DATA_BLOCK "DB_ALARM"   // DB100
{ S7_Optimized_Access := 'FALSE' }
VERSION : 0.1
   VAR
      ALARM : Struct
         ALARM_GLOBAL : Bool;   // globální alarm
         HERMA_ERROR : Bool;
         ALARM_2 : Bool;
         ALARM_3 : Bool;
         ALARM_4 : Bool;
         ALARM_5 : Bool;
         air : Bool;   // nedostatečný tlak vzduchu
         ALARM_7 : Bool;
         ALARM_8 : Bool;
         ALARM_9 : Bool;
         ALARM_10 : Bool;
         ALARM_11 : Bool;
         ALARM_12 : Bool;
         ALARM_13 : Bool;
         ALARM_14 : Bool;
         vypadek_safety_karty : Bool;
      END_STRUCT;
      WRONG : Struct
         NENI_INICIALIZACE : Bool;
         WRONG_global : Bool;
         dvere_L_tevreny : Bool;
         dvere_P_otevreny : Bool;
         WRONG_4 : Bool;
         WRONG_5 : Bool;
         WRONG_6 : Bool;
         WRONG_7 : Bool;
         WRONG_8 : Bool;
         WRONG_9 : Bool;
         WRONG_10 : Bool;
         WRONG_11 : Bool;
         WRONG_12 : Bool;
         WRONG_13 : Bool;
         rop_glob_warning : Bool;
         rop_active_autocale : Bool;
      END_STRUCT;
      OP0 : Struct
         ALARM : Struct
            DOOR_ERROR : Bool;
            ALARM_1 : Bool;
            ALARM_2 : Bool;
            ALARM_3 : Bool;
            ALARM_4 : Bool;
            ALARM_5 : Bool;
            ALARM_6 : Bool;
            ALARM_7 : Bool;
            ALARM_8 : Bool;
            ALARM_9 : Bool;
            ALARM_10 : Bool;
            ALARM_11 : Bool;
            ALARM_12 : Bool;
            ALARM_13 : Bool;
            ALARM_14 : Bool;
            ALARM_15 : Bool;
         END_STRUCT;
         WRONG : Struct
            WRONG_0 : Bool;
            WRONG_1 : Bool;
            WRONG_2 : Bool;
            WRONG_3 : Bool;
            WRONG_4 : Bool;
            WRONG_5 : Bool;
            WRONG_6 : Bool;
            WRONG_7 : Bool;
            WRONG_8 : Bool;
            WRONG_9 : Bool;
            WRONG_10 : Bool;
            WRONG_11 : Bool;
            WRONG_12 : Bool;
            WRONG_13 : Bool;
            WRONG_14 : Bool;
            WRONG_15 : Bool;
         END_STRUCT;
         M_0 : Int;
         M_1 : Int;
         M_2 : Int;
         M_3 : Int;
         M_4 : Int;
         M_5 : Int;
         M_6 : Int;
         M_7 : Int;
         M_8 : Int;
         M_9 : Int;
         M_10 : Int;
         M_11 : Int;
         M_12 : Int;
         M_13 : Int;
         M_14 : Int;
         M_15 : Int;
      END_STRUCT;
      OP1 : Struct
         ALARM : Struct
            dvere_1 : Bool;
            ALARM_1 : Bool;
            ALARM_2 : Bool;
            ALARM_3 : Bool;
            ALARM_4 : Bool;
            ALARM_5 : Bool;
            ALARM_6 : Bool;
            hladina_mimo_mez : Bool;
            ALARM_8 : Bool;
            ALARM_9 : Bool;
            ALARM_10 : Bool;
            ALARM_11 : Bool;
            ALARM_12 : Bool;
            ALARM_13 : Bool;
            ALARM_14 : Bool;
            ALARM_15 : Bool;
         END_STRUCT;
         WRONG : Struct
            WRONG_0 : Bool;
            WRONG_1 : Bool;
            WRONG_2 : Bool;
            WRONG_3 : Bool;
            WRONG_4 : Bool;
            WRONG_5 : Bool;
            WRONG_6 : Bool;
            WRONG_7 : Bool;
            WRONG_8 : Bool;
            WRONG_9 : Bool;
            WRONG_10 : Bool;
            WRONG_11 : Bool;
            WRONG_12 : Bool;
            WRONG_13 : Bool;
            WRONG_14 : Bool;
            WRONG_15 : Bool;
         END_STRUCT;
         "-Y7_KARUSEL" : Int;
         "-Y9_ZARAZKA" : Int;
         M_2 : Int;
         M_3 : Int;
         M_4 : Int;
         M_5 : Int;
         M_6 : Int;
         M_7 : Int;
         M_8 : Int;
         M_9 : Int;
         M_10 : Int;
         M_11 : Int;
         M_12 : Int;
         M_13 : Int;
         M_14 : Int;
         M_15 : Int;
      END_STRUCT;
      OP2 : Struct
         ALARM : Struct
            dvere_1 : Bool;
            dvere_2 : Bool;
            dvere_3 : Bool;
            dvere_4 : Bool;
            paprsek : Bool;
            porucha_svarovani : Bool;
            rop_alarm : Bool;
            servo_power_error : Bool;
            servo_jog_error : Bool;
            servo_homing : Bool;
            Cel_podel_porucha : Bool;
            vysoka_tuzka : Bool;
            ALARM_12 : Bool;
            ALARM_13 : Bool;
            folie : Bool;
            ALARM_15 : Bool;
         END_STRUCT;
         WRONG : Struct
            WRONG_0 : Bool;
            WRONG_1 : Bool;
            WRONG_2 : Bool;
            WRONG_3 : Bool;
            WRONG_4 : Bool;
            WRONG_5 : Bool;
            WRONG_6 : Bool;
            WRONG_7 : Bool;
            WRONG_8 : Bool;
            WRONG_9 : Bool;
            WRONG_10 : Bool;
            WRONG_11 : Bool;
            WRONG_12 : Bool;
            WRONG_13 : Bool;
            WRONG_14 : Bool;
            WRONG_15 : Bool;
         END_STRUCT;
         A1 : Int;   // -YA1
         A2 : Int;   // -YA2
         A3 : Int;   // -YA3
         A4 : Int;   // -YA4
         A5 : Int;   // -YA5
         A6 : Int;   // -YA6
         A7 : Int;   // -YA7
         A8 : Int;   // -YA8
         M_8 : Int;
         M_9 : Int;
         M_10 : Int;
         M_11 : Int;
         M_12 : Int;
         M_13 : Int;
         M_14 : Int;
         M_15 : Int;
      END_STRUCT;
      OP3 : Struct
         ALARM : Struct
            ALARM_0 : Bool;
            ALARM_1 : Bool;
            ALARM_2 : Bool;
            ALARM_3 : Bool;
            ALARM_4 : Bool;
            ALARM_5 : Bool;
            ALARM_6 : Bool;
            ALARM_7 : Bool;
            ALARM_8 : Bool;
            ALARM_9 : Bool;
            ALARM_10 : Bool;
            ALARM_11 : Bool;
            ALARM_12 : Bool;
            ALARM_13 : Bool;
            ALARM_14 : Bool;
            ALARM_15 : Bool;
         END_STRUCT;
         WRONG : Struct
            WRONG_0 : Bool;
            WRONG_1 : Bool;
            WRONG_2 : Bool;
            WRONG_3 : Bool;
            WRONG_4 : Bool;
            WRONG_5 : Bool;
            WRONG_6 : Bool;
            WRONG_7 : Bool;
            WRONG_8 : Bool;
            WRONG_9 : Bool;
            WRONG_10 : Bool;
            WRONG_11 : Bool;
            WRONG_12 : Bool;
            WRONG_13 : Bool;
            WRONG_14 : Bool;
            WRONG_15 : Bool;
         END_STRUCT;
         B1 : Int;   // -YB1
         B2 : Int;   // -YB2
         B3 : Int;   // -YB3
         B4 : Int;   // -YB4
         B5 : Int;   // -YB5
         B6 : Int;   // -YB6
         B7 : Int;   // -YB7
         B8 : Int;   // -YB8
         M_8 : Int;
         M_9 : Int;
         M_10 : Int;
         M_11 : Int;
         M_12 : Int;
         M_13 : Int;
         M_14 : Int;
         M_15 : Int;
      END_STRUCT;
      OP4 : Struct
         ALARM : Struct
            odsavani_nefunguje : Bool;
            ALARM_1 : Bool;
            ALARM_2 : Bool;
            ALARM_3 : Bool;
            ALARM_4 : Bool;
            ALARM_5 : Bool;
            ALARM_6 : Bool;
            ALARM_7 : Bool;
            ALARM_8 : Bool;
            ALARM_9 : Bool;
            ALARM_10 : Bool;
            ALARM_11 : Bool;
            ALARM_12 : Bool;
            ALARM_13 : Bool;
            ALARM_14 : Bool;
            ALARM_15 : Bool;
         END_STRUCT;
         WRONG : Struct
            WRONG_0 : Bool;
            WRONG_1 : Bool;
            WRONG_2 : Bool;
            WRONG_3 : Bool;
            WRONG_4 : Bool;
            WRONG_5 : Bool;
            WRONG_6 : Bool;
            WRONG_7 : Bool;
            WRONG_8 : Bool;
            WRONG_9 : Bool;
            WRONG_10 : Bool;
            WRONG_11 : Bool;
            WRONG_12 : Bool;
            WRONG_13 : Bool;
            WRONG_14 : Bool;
            WRONG_15 : Bool;
         END_STRUCT;
         M_0 : Int;
         M_1 : Int;
         M_2 : Int;
         M_3 : Int;
         M_4 : Int;
         M_5 : Int;
         M_6 : Int;
         M_7 : Int;
         M_8 : Int;
         M_9 : Int;
         M_10 : Int;
         M_11 : Int;
         M_12 : Int;
         M_13 : Int;
         M_14 : Int;
         M_15 : Int;
      END_STRUCT;
      OP5 : Struct
         ALARM : Struct
            ALARM_0 : Bool;
            ALARM_1 : Bool;
            ALARM_2 : Bool;
            ALARM_3 : Bool;
            ALARM_4 : Bool;
            ALARM_5 : Bool;
            ALARM_6 : Bool;
            ALARM_7 : Bool;
            ALARM_8 : Bool;
            ALARM_9 : Bool;
            ALARM_10 : Bool;
            ALARM_11 : Bool;
            ALARM_12 : Bool;
            ALARM_13 : Bool;
            ALARM_14 : Bool;
            ALARM_15 : Bool;
         END_STRUCT;
         WRONG : Struct
            WRONG_0 : Bool;
            WRONG_1 : Bool;
            WRONG_2 : Bool;
            WRONG_3 : Bool;
            WRONG_4 : Bool;
            WRONG_5 : Bool;
            WRONG_6 : Bool;
            WRONG_7 : Bool;
            WRONG_8 : Bool;
            WRONG_9 : Bool;
            WRONG_10 : Bool;
            WRONG_11 : Bool;
            WRONG_12 : Bool;
            WRONG_13 : Bool;
            WRONG_14 : Bool;
            WRONG_15 : Bool;
         END_STRUCT;
         M_0 : Int;
         M_1 : Int;
         M_2 : Int;
         M_3 : Int;
         M_4 : Int;
         M_5 : Int;
         M_6 : Int;
         M_7 : Int;
         M_8 : Int;
         M_9 : Int;
         M_10 : Int;
         M_11 : Int;
         M_12 : Int;
         M_13 : Int;
         M_14 : Int;
         M_15 : Int;
      END_STRUCT;
      null : Struct
         ALARM_0 : Bool;
         ALARM_1 : Bool;
         ALARM_2 : Bool;
         ALARM_3 : Bool;
         ALARM_4 : Bool;
         ALARM_5 : Bool;
         ALARM_6 : Bool;
         ALARM_7 : Bool;
         ALARM_8 : Bool;
         ALARM_9 : Bool;
         ALARM_10 : Bool;
         ALARM_11 : Bool;
         ALARM_12 : Bool;
         ALARM_13 : Bool;
         ALARM_14 : Bool;
         ALARM_15 : Bool;
      END_STRUCT;
      alarmy : Array[0..255] of Bool;
      alarm_line : Int;
      wrong_line : Int;
      alarm_op_1 : Int;
      wrong_op_1 : Int;
      alarm_op_2 : Int;
      wrong_op_2 : Int;
      alarm_op_3 : Int;
      wrong_op_3 : Int;
      alarm_op_4 : Int;
      wrong_op_4 : Int;
      alarm_op_5 : Int;
      wrong_op_5 : Int;
      T_tiskarna : TON_TIME;
   END_VAR
BEGIN
END_DATA_BLOCK

// folder: STANDARD/BLOKY_DO_OPERACI

DATA_BLOCK "DB_STS_M"   // DB101
{ S7_Optimized_Access := 'FALSE' }
VERSION : 0.1
   VAR
      OP0 : Struct
         STS_M0 : UInt;
         STS_M1 : UInt;
         STS_M2 : UInt;
         STS_M3 : UInt;
         STS_M4 : UInt;
         STS_M5 : UInt;
         STS_M6 : UInt;
         STS_M7 : UInt;
         STS_M8 : UInt;
         STS_M9 : UInt;
         STS_M10 : UInt;
         STS_M11 : UInt;
         STS_M12 : UInt;
         STS_M13 : UInt;
         STS_M14 : UInt;
         STS_M15 : UInt;
      END_STRUCT;
      OP1 : Struct
         KARUSEL : UInt;
         ZARAZKA : UInt;
         STS_M2 : UInt;
         STS_M3 : UInt;
         STS_M4 : UInt;
         STS_M5 : UInt;
         STS_M6 : UInt;
         STS_M7 : UInt;
         STS_M8 : UInt;
         STS_M9 : UInt;
         STS_M10 : UInt;
         STS_M11 : UInt;
         STS_M12 : UInt;
         STS_M13 : UInt;
         STS_M14 : UInt;
         STS_M15 : UInt;
         OP1 : Struct
            STS_M0 : UInt;
            STS_M1 : UInt;
            STS_M2 : UInt;
            STS_M3 : UInt;
            STS_M4 : UInt;
            STS_M5 : UInt;
            STS_M6 : UInt;
            STS_M7 : UInt;
            STS_M8 : UInt;
            STS_M9 : UInt;
            STS_M10 : UInt;
            STS_M11 : UInt;
            STS_M12 : UInt;
            STS_M13 : UInt;
            STS_M14 : UInt;
            STS_M15 : UInt;
         END_STRUCT;
      END_STRUCT;
      OP2 : Struct
         A1 : UInt;
         A2 : UInt;
         A3 : UInt;
         A4 : UInt;
         A5 : UInt;
         A6 : UInt;
         A7 : UInt;
         A8 : UInt;
         STS_M8 : UInt;
         STS_M9 : UInt;
         STS_M10 : UInt;
         STS_M11 : UInt;
         STS_M12 : UInt;
         STS_M13 : UInt;
         STS_M14 : UInt;
         STS_M15 : UInt;
      END_STRUCT;
      OP3 : Struct
         B1 : UInt;
         B2 : UInt;
         B3 : UInt;
         B4 : UInt;
         B5 : UInt;
         B6 : UInt;
         B7 : UInt;
         B8 : UInt;
         STS_M8 : UInt;
         STS_M9 : UInt;
         STS_M10 : UInt;
         STS_M11 : UInt;
         STS_M12 : UInt;
         STS_M13 : UInt;
         STS_M14 : UInt;
         STS_M15 : UInt;
      END_STRUCT;
   END_VAR
BEGIN
END_DATA_BLOCK

// folder: STANDARD/CORE/FB_ABMARK_PROFINET

DATA_BLOCK "OVLADANI_LASER_DB"   // DB400
{ S7_Optimized_Access := 'TRUE' }
VERSION : 0.1
// stored: InstanceOfName OVLADANI_LASER
"OVLADANI_LASER"
BEGIN
END_DATA_BLOCK

DATA_BLOCK "DB_DATA_LASER"   // DB401
{ S7_Optimized_Access := 'TRUE' }
VERSION : 0.1
   VAR
      LASER_DATA_READ : Array[0..71] of Byte;
      LASER_DATA_WRITE : Array[0..71] of Byte;
      READ : Bool;
      WRITE : Bool;
   END_VAR
BEGIN
END_DATA_BLOCK

DATA_BLOCK "DB_LASER"   // DB402
{ S7_Optimized_Access := 'TRUE' }
VERSION : 0.1
   VAR
      DATA_DO_ETIKETY : Struct
         TEXT : String[5];
         "INT" : Int;
         "REAL" : Real;
         PROGRAM : Array[0..1] of String[10];
      END_STRUCT;
      DATA_DO_DAT : Struct
         ZAVORKA_L : Char := '<';
         ZAVORKA_P : Char := '>';
         XLP : Array[0..3] of Char;
      END_STRUCT;
      smaz_me_start : Bool;
      smaz_me_adresa : Int;
   END_VAR
BEGIN
   DATA_DO_DAT.XLP[0] := '.';
   DATA_DO_DAT.XLP[1] := 'x';
   DATA_DO_DAT.XLP[2] := 'l';
   DATA_DO_DAT.XLP[3] := 'p';
   DATA_DO_ETIKETY.PROGRAM[0] := 'TEST_1';
   DATA_DO_ETIKETY.PROGRAM[1] := 'TEST_222';
END_DATA_BLOCK

// folder: STANDARD/LINE

DATA_BLOCK "CONTROL_LINE_DB"   // DB27
{ S7_Optimized_Access := 'TRUE' }
VERSION : 0.1
// stored: InstanceOfName CONTROL_LINE
"CONTROL_LINE"
BEGIN
END_DATA_BLOCK

// folder: System blocks/Program resources

DATA_BLOCK "A3-PLC1214_Connection_DB"   // DB5
{ S7_Optimized_Access := 'TRUE' }
AUTHOR : SIMATIC
FAMILY : MC7Plus
NAME : TC_IP_v4
VERSION : 1.0
// stored: InstanceOfName TCON_IP_v4
"TCON_IP_v4"
BEGIN
   ID := 1;
   InterfaceId := 64;
   RemotePort := 25001;
   ActiveEstablished := true;
   RemoteAddress.ADDR[1] := 192;
   RemoteAddress.ADDR[2] := 168;
   RemoteAddress.ADDR[4] := 100;
END_DATA_BLOCK

// folder: (top level)

ORGANIZATION_BLOCK "Main"   // OB1, LAD, ProgramCycle
TITLE = "Main Program Sweep (Cycle)"
{ S7_Optimized_Access := 'TRUE' }
VERSION : 0.1
   VAR_INPUT
      Initial_Call : Bool;   // Initial call of this OB
      Remanence : Bool;   // =True, if remanent data are available
   END_VAR
BEGIN

REGION Network 1
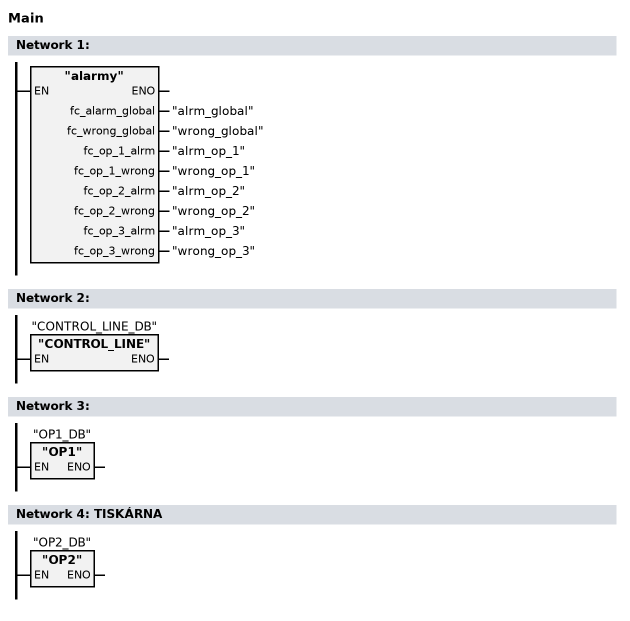
   RUNG wire#powerrail
      "alarmy"(fc_alarm_global => "alrm_global", fc_wrong_global => "wrong_global", fc_op_1_alrm => "alrm_op_1", fc_op_1_wrong => "wrong_op_1", fc_op_2_alrm => "alrm_op_2", fc_op_2_wrong => "wrong_op_2", fc_op_3_alrm => "alrm_op_3", fc_op_3_wrong => "wrong_op_3")
   END_RUNG
   // the same network as SCL:
   "alarmy"(fc_alarm_global => "alrm_global",
            fc_wrong_global => "wrong_global",
            fc_op_1_alrm => "alrm_op_1",
            fc_op_1_wrong => "wrong_op_1",
            fc_op_2_alrm => "alrm_op_2",
            fc_op_2_wrong => "wrong_op_2",
            fc_op_3_alrm => "alrm_op_3",
            fc_op_3_wrong => "wrong_op_3");
END_REGION

REGION Network 2
   RUNG wire#powerrail
      "CONTROL_LINE_DB"()
   END_RUNG
   // the same network as SCL:
   "CONTROL_LINE_DB"();   // "CONTROL_LINE"
END_REGION

REGION Network 3
   RUNG wire#powerrail
      "OP1_DB"()
   END_RUNG
   // the same network as SCL:
   "OP1_DB"();   // "OP1"
END_REGION

REGION Network 4: TISKÁRNA
   RUNG wire#powerrail
      "OP2_DB"()
   END_RUNG
   // the same network as SCL:
   "OP2_DB"();   // "OP2"
END_REGION
END_ORGANIZATION_BLOCK

ORGANIZATION_BLOCK "CyclicInterrupt"   // OB30, LAD, CyclicInterrupt
{ S7_Optimized_Access := 'TRUE' }
VERSION : 0.1
   VAR_INPUT
      Initial_Call : Bool;   // Initial call of this OB
      Event_Count : Int;   // Events discarded
   END_VAR
   VAR_TEMP
      AKTUALNI_POZICE_FOLIE : DInt;
      AKTUALNI_POZICE_ETIKETA : DInt;
   END_VAR
   VAR_TEMP   // added for the SCL form of the ladder/FBD networks
      _w1 : Bool;
   END_VAR
BEGIN

REGION Network 1
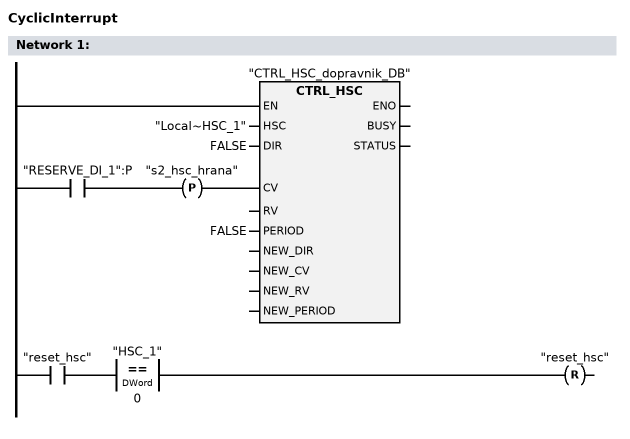
   #_w1 := "RESERVE_DI_1":P AND NOT "s2_hsc_hrana";   // rising edge
   "s2_hsc_hrana" := "RESERVE_DI_1":P;
   "CTRL_HSC_dopravnik_DB"(HSC := "Local~HSC_1", DIR := FALSE, CV := #_w1, PERIOD := FALSE);   // CTRL_HSC
   IF "reset_hsc" AND ("HSC_1" = 0) THEN "reset_hsc" := FALSE; END_IF;
END_REGION

REGION Network 2 (SCL): Poloha plata od s2 [mm]
   // aktualni_poloha = HSC_1 × mm/puls (fourfold). HSC se nuluje na náběhu s2 (síť 1).
   // Konstanta 1.488 = mm na 1 puls – LIMIT brání přetečení při chodu naprázdno.
   "DB_HMI_recype".aktualni_poloha := REAL_TO_DINT(LIMIT(MN := 0.0,
                                                                                                         IN := DINT_TO_REAL(DWORD_TO_DINT("HSC_1":P)) * 4,
                                                                                                         MX := 99999.0));
END_REGION
END_ORGANIZATION_BLOCK

// folder: OPERACE

FUNCTION_BLOCK "OP0"   // FB49, LAD
{ S7_Optimized_Access := 'TRUE' }
VERSION : 0.1
   VAR
      CONTROL_MAN : Struct
         B0 : Bool;
         B1 : Bool;
         B2 : Bool;
         B3 : Bool;
         B4 : Bool;
         B5 : Bool;
         B6 : Bool;
         B7 : Bool;
         B8 : Bool;
         B9 : Bool;
         B10 : Bool;
         B11 : Bool;
         B12 : Bool;
         B13 : Bool;
         B14 : Bool;
         B15 : Bool;
         B16 : Bool;
         B17 : Bool;
         B18 : Bool;
         B19 : Bool;
         B20 : Bool;
         B21 : Bool;
         B22 : Bool;
         B23 : Bool;
         B24 : Bool;
         B25 : Bool;
         B26 : Bool;
         B27 : Bool;
         B28 : Bool;
         B29 : Bool;
         B30 : Bool;
         B31 : Bool;
      END_STRUCT;
      CONTROL_AUTOMAT : Struct
         B0 : Bool;
         B1 : Bool;
         B2 : Bool;
         B3 : Bool;
         B4 : Bool;
         B5 : Bool;
         B6 : Bool;
         B7 : Bool;
         B8 : Bool;
         B9 : Bool;
         B10 : Bool;
         B11 : Bool;
         B12 : Bool;
         B13 : Bool;
         B14 : Bool;
         B15 : Bool;
         B16 : Bool;
         B17 : Bool;
         B18 : Bool;
         B19 : Bool;
         B20 : Bool;
         B21 : Bool;
         B22 : Bool;
         B23 : Bool;
         B24 : Bool;
         B25 : Bool;
         B26 : Bool;
         B27 : Bool;
         B28 : Bool;
         B29 : Bool;
         B30 : Bool;
         B31 : Bool;
      END_STRUCT;
      SENSORS : Struct
         S0 : Bool;
         S1 : Bool;
         S2 : Bool;
         S3 : Bool;
         S4 : Bool;
         S5 : Bool;
         S6 : Bool;
         S7 : Bool;
         S8 : Bool;
         S9 : Bool;
         S10 : Bool;
         S11 : Bool;
         S12 : Bool;
         S13 : Bool;
         S14 : Bool;
         S15 : Bool;
         S16 : Bool;
         S17 : Bool;
         S18 : Bool;
         S19 : Bool;
         S20 : Bool;
         S21 : Bool;
         S22 : Bool;
         S23 : Bool;
         S24 : Bool;
         S25 : Bool;
         S26 : Bool;
         S27 : Bool;
         S28 : Bool;
         S29 : Bool;
         S30 : Bool;
         S31 : Bool;
      END_STRUCT;
      SENSORS_1 : Struct
         S0 : Bool;
         S1 : Bool;
         S2 : Bool;
         S3 : Bool;
         S4 : Bool;
         S5 : Bool;
         S6 : Bool;
         S7 : Bool;
         S8 : Bool;
         S9 : Bool;
         S10 : Bool;
         S11 : Bool;
         S12 : Bool;
         S13 : Bool;
         S14 : Bool;
         S15 : Bool;
         S16 : Bool;
         S17 : Bool;
         S18 : Bool;
         S19 : Bool;
         S20 : Bool;
         S21 : Bool;
         S22 : Bool;
         S23 : Bool;
         S24 : Bool;
         S25 : Bool;
         S26 : Bool;
         S27 : Bool;
         S28 : Bool;
         S29 : Bool;
         S30 : Bool;
         S31 : Bool;
      END_STRUCT;
      S_0 : "SENSOR";
      S_1 : "SENSOR";
      S_2 : "SENSOR";
      S_3 : "SENSOR";
      S_4 : "SENSOR";
      S_5 : "SENSOR";
      S_6 : "SENSOR";
      S_7 : "SENSOR";
      S_8 : "SENSOR";
      S_9 : "SENSOR";
      s_10 : "SENSOR";
      S_11 : "SENSOR";
      S_12 : "SENSOR";
      S_13 : "SENSOR";
      S_14 : "SENSOR";
      S_15 : "SENSOR";
      S_16 : "SENSOR";
      S_17 : "SENSOR";
      S_18 : "SENSOR";
      S_19 : "SENSOR";
      S_20 : "SENSOR";
      S_21 : "SENSOR";
      S_22 : "SENSOR";
      S_23 : "SENSOR";
      S_24 : "SENSOR";
      S_25 : "SENSOR";
      S_26 : "SENSOR";
      S_27 : "SENSOR";
      S_28 : "SENSOR";
      S_29 : "SENSOR";
      S_30 : "SENSOR";
      S_31 : "SENSOR";
      S_32 : "SENSOR";
      S_33 : "SENSOR";
      S_34 : "SENSOR";
      S_35 : "SENSOR";
      M_0 : "MOTOR_CONTROL_BLOCK";
      M_1 : "MOTOR_CONTROL_BLOCK";
      M_2 : "MOTOR_CONTROL_BLOCK";
      M_3 : "MOTOR_CONTROL_BLOCK";
      SQCR : Int;
      TRIG : Struct
         inicial_ok_op : Bool;
         DSSAD : Bool;
         INICIALIZACE_PROBEHLA : Bool;
         trig_dil : Bool;
         p_trig_control_tcon : Bool;
         T6 : Bool;
         T7 : Bool;
         T8 : Bool;
         T9 : Bool;
         T10 : Bool;
         T11 : Bool;
         T12 : Bool;
         T13 : Bool;
         T14 : Bool;
         T15 : Bool;
         T16 : Bool;
         T17 : Bool;
      END_STRUCT;
      MEMOR : Struct
         M0 : Bool;
         M1 : Bool;
         M2 : Bool;
         M3 : Bool;
         M4 : Bool;
         M5 : Bool;
         M6 : Bool;
         M7 : Bool;
         M8 : Bool;
         M9 : Bool;
         M10 : Bool;
         M11 : Bool;
         RESET_ERROR : Bool;
         M13 : Bool;
         M14 : Bool;
         M15 : Bool;
         M16 : Bool;
         M17 : Bool;
         M18 : Bool;
         M19 : Bool;
         M20 : Bool;
         M21 : Bool;
         M22 : Bool;
         M23 : Bool;
         M24 : Bool;
         M25 : Bool;
         M26 : Bool;
         M27 : Bool;
         M28 : Bool;
         M29 : Bool;
         M30 : Bool;
         M31 : Bool;
         M32 : Bool;
         M33 : Bool;
         start_caklu : Bool;
         M35 : Bool;
         M36 : Bool;
         M37 : Bool;
         M38 : Bool;
         M39 : Bool;
         ALARM_GLOBAL : Bool;
         M41 : Bool;
         M42 : Bool;
         M43 : Bool;
         M44 : Bool;
         M45 : Bool;
         M46 : Bool;
         M47 : Bool;
         M48 : Bool;
         M49 : Bool;
         M50 : Bool;
         M51 : Bool;
         M52 : Bool;
         M53 : Bool;
         M54 : Bool;
         M55 : Bool;
         M56 : Bool;
         M57 : Bool;
         M58 : Bool;
         M59 : Bool;
         M60 : Bool;
         M61 : Bool;
         M62 : Bool;
         M63 : Bool;
      END_STRUCT;
      "TIMER" : Struct
         TIMER_0 : IEC_TIMER;
         TIMER_VACUUM_CLEANER : IEC_TIMER;
         TIMER_DELAY_RESET_EXECUTE : IEC_TIMER;
         TIMER_3 : IEC_TIMER;
         TIMER_4 : IEC_TIMER;
         TIMER_5 : IEC_TIMER;
         TIMER_6 : IEC_TIMER;
         TIMER_7 : IEC_TIMER;
      END_STRUCT;
      HMI : Struct
         povoleni_volby_receptu : Bool;
         "svetlo_on/off" : Bool;
         ALARM_VIDITELNOST : Bool;
         hmi_3 : Bool;
         hmi_4 : Bool;
         hmi_5 : Bool;
         hmi_6 : Bool;
         hmi_7 : Bool;
         hmi_8 : Bool;
         hmi_9 : Bool;
         hmi_10 : Bool;
         hmi_11 : Bool;
         hmi_12 : Bool;
         hmi_13 : Bool;
         hmi_14 : Bool;
         hmi_15 : Bool;
      END_STRUCT;
      kontrola_tcon : Int;
      cyklus_aretace : Int;
      string_pam : String;
      error_m1 : Int;
      error_m2 : Int;
      MAXA : Struct
         ACTUAL_MESSAGE : String[16];
         name_char : Array[0..16] of Char;
         adresace : Byte;
      END_STRUCT;
      HMI_SPEED : Real;
      hmi_man_cab : Bool;
      HMI_START : Bool;
      TRIGR_LASER : DWord;
   END_VAR
   VAR_TEMP
      DATA : Array[0..255] of Char;
      PREVOD : Int;
      NORM_SCALE : LReal;
   END_VAR
   VAR CONSTANT
      STEP_0 : Int := 0;
      step_2 : Int := 2;
      STEP_4 : Int := 4;
      STEP_5_HOME : Int := 5;
      STEP_7 : Int := 7;
      STEP_10 : Int := 10;
      STEP_15 : Int := 15;
      STEP_20 : Int := 20;
      STEP_23 : Int := 23;
      STEP_25 : Int := 25;
      STEP_27 : Int := 27;
      STEP_30 : Int := 30;
      STEP_35 : Int := 35;
      STEP_37 : Int := 37;
      STEP_40 : Int := 40;
      STEP_45 : Int := 45;
      STEP_50 : Int := 50;
      STEP_55 : Int := 55;
      STEP_60 : Int := 60;
      STEP_65 : Int := 65;
      STEP_70 : Int := 70;
      STEP_75 : Int := 75;
      STEP_80 : Int := 80;
      STEP_83 : Int := 83;
      STEP_85 : Int := 85;
      STEP_90 : Int := 90;
      STEP_95 : Int := 95;
      STEP_100 : Int := 100;
      STEP_105 : Int := 105;
      STEP_110 : Int := 110;
      STEP_113 : Int := 113;
      STEP_115 : Int := 115;
      STEP_120 : Int := 120;
      STEP_125 : Int := 125;
      STEP_130 : Int := 130;
      STEP_135 : Int := 135;
      STEP_140 : Int := 140;
      STEP_145 : Int := 145;
      STEP_150 : Int := 150;
      STEP_155 : Int := 155;
      STEP_1000_KONTROLA : Int := 1000;
      STEP_1005_START_INICIAL : Int := 1005;
      STEP_1010_close_door : Int := 1010;
      STEP_1015 : Int := 1015;
      STEP_1020_HOME_OK : Int := 1020;
      STEP_1025 : Int := 1025;
      STEP_3000 : Int := 3000;
      STEP_3005 : Int := 3005;
      STEP_3010 : Int := 3010;
      STEP_3015 : Int := 3015;
      STEP_3020 : Int := 3020;
      STEP_2000 : Int := 2000;
      string_null : String;
      char_null : Char;
   END_VAR
   VAR_TEMP   // added for the SCL form of the ladder/FBD networks
      _w1 : Bool;
      _w2 : Bool;
      _w3 : Bool;
      _w4 : Bool;
      _w5 : Bool;
      _w6 : Bool;
      _w7 : Bool;
      _w8 : Bool;
      _w9 : Bool;
   END_VAR
BEGIN

REGION Network 1 (SCL)
   IF "FirstScan" = true THEN
       #MAXA.adresace := 0;
   END_IF;
     (*  

   #MAXA.name_char[0] := "-XT500_name_byte_0";
   #MAXA.name_char[1] := "-XT500_name_byte_1";
   #MAXA.name_char[2] := "-XT500_name_byte_2";
   #MAXA.name_char[3] := "-XT500_name_byte_3";
   #MAXA.name_char[4] := "-XT500_name_byte_4";
   #MAXA.name_char[5] := "-XT500_name_byte_5";
   #MAXA.name_char[6] := "-XT500_name_byte_6";
   #MAXA.name_char[7] := "-XT500_name_byte_7";
   #MAXA.name_char[8] := "-XT500_name_byte_8";
   #MAXA.name_char[9] := "-XT500_name_byte_9";
   #MAXA.name_char[10] := "-XT500_name_byte_10";
   #MAXA.name_char[11] := "-XT500_name_byte_11";
   #MAXA.name_char[12] := "-XT500_name_byte_12";
   #MAXA.name_char[13] := "-XT500_name_byte_13";
   #MAXA.name_char[14] := "-XT500_name_byte_14";
   #MAXA.name_char[15] := "-XT500_name_byte_15";
   *)

   IF #SQCR <> 0 THEN
       IF #MAXA.adresace > 16 THEN
           #MAXA.adresace := 0;
       END_IF;
       #MAXA.ACTUAL_MESSAGE[#MAXA.adresace + 1] := #MAXA.name_char[#MAXA.adresace];
       #MAXA.adresace := #MAXA.adresace + 1;
   END_IF;
END_REGION

REGION Network 2: manuali ovladani reset
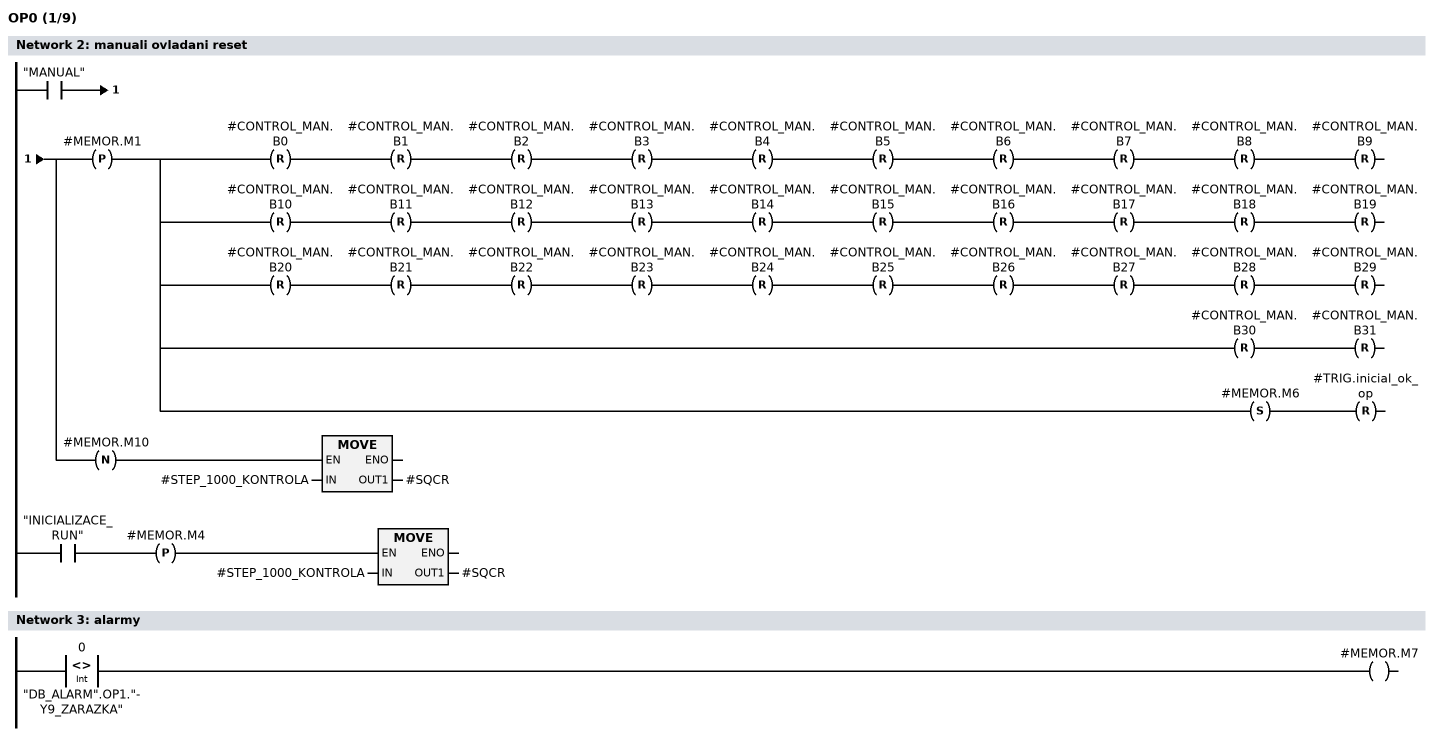
   RUNG wire#powerrail
      Contact( "MANUAL" )
      wire#w1
      P_Trig( #MEMOR.M1 )
      wire#w2
      R_Coil( #CONTROL_MAN.B0 )
      R_Coil( #CONTROL_MAN.B1 )
      R_Coil( #CONTROL_MAN.B2 )
      R_Coil( #CONTROL_MAN.B3 )
      R_Coil( #CONTROL_MAN.B4 )
      R_Coil( #CONTROL_MAN.B5 )
      R_Coil( #CONTROL_MAN.B6 )
      R_Coil( #CONTROL_MAN.B7 )
      R_Coil( #CONTROL_MAN.B8 )
      R_Coil( #CONTROL_MAN.B9 )
   END_RUNG
   RUNG wire#w2
      R_Coil( #CONTROL_MAN.B10 )
      R_Coil( #CONTROL_MAN.B11 )
      R_Coil( #CONTROL_MAN.B12 )
      R_Coil( #CONTROL_MAN.B13 )
      R_Coil( #CONTROL_MAN.B14 )
      R_Coil( #CONTROL_MAN.B15 )
      R_Coil( #CONTROL_MAN.B16 )
      R_Coil( #CONTROL_MAN.B17 )
      R_Coil( #CONTROL_MAN.B18 )
      R_Coil( #CONTROL_MAN.B19 )
   END_RUNG
   RUNG wire#w2
      R_Coil( #CONTROL_MAN.B20 )
      R_Coil( #CONTROL_MAN.B21 )
      R_Coil( #CONTROL_MAN.B22 )
      R_Coil( #CONTROL_MAN.B23 )
      R_Coil( #CONTROL_MAN.B24 )
      R_Coil( #CONTROL_MAN.B25 )
      R_Coil( #CONTROL_MAN.B26 )
      R_Coil( #CONTROL_MAN.B27 )
      R_Coil( #CONTROL_MAN.B28 )
      R_Coil( #CONTROL_MAN.B29 )
   END_RUNG
   RUNG wire#w2
      R_Coil( #CONTROL_MAN.B30 )
      R_Coil( #CONTROL_MAN.B31 )
   END_RUNG
   RUNG wire#w2
      S_Coil( #MEMOR.M6 )
      R_Coil( #TRIG.inicial_ok_op )
   END_RUNG
   RUNG wire#w1
      N_Trig( #MEMOR.M10 )
      Move(in := #STEP_1000_KONTROLA, out1 => #SQCR)
   END_RUNG
   RUNG wire#powerrail
      Contact( "INICIALIZACE_RUN" )
      P_Trig( #MEMOR.M4 )
      Move(in := #STEP_1000_KONTROLA, out1 => #SQCR)
   END_RUNG
   // the same network as SCL:
   #_w1 := "MANUAL" AND NOT #MEMOR.M1;   // rising edge
   #MEMOR.M1 := "MANUAL";
   IF #_w1 THEN
       #CONTROL_MAN.B0 := FALSE;
       #CONTROL_MAN.B1 := FALSE;
       #CONTROL_MAN.B2 := FALSE;
       #CONTROL_MAN.B3 := FALSE;
       #CONTROL_MAN.B4 := FALSE;
       #CONTROL_MAN.B5 := FALSE;
       #CONTROL_MAN.B6 := FALSE;
       #CONTROL_MAN.B7 := FALSE;
       #CONTROL_MAN.B8 := FALSE;
       #CONTROL_MAN.B9 := FALSE;
       #CONTROL_MAN.B10 := FALSE;
       #CONTROL_MAN.B11 := FALSE;
       #CONTROL_MAN.B12 := FALSE;
       #CONTROL_MAN.B13 := FALSE;
       #CONTROL_MAN.B14 := FALSE;
       #CONTROL_MAN.B15 := FALSE;
       #CONTROL_MAN.B16 := FALSE;
       #CONTROL_MAN.B17 := FALSE;
       #CONTROL_MAN.B18 := FALSE;
       #CONTROL_MAN.B19 := FALSE;
       #CONTROL_MAN.B20 := FALSE;
       #CONTROL_MAN.B21 := FALSE;
       #CONTROL_MAN.B22 := FALSE;
       #CONTROL_MAN.B23 := FALSE;
       #CONTROL_MAN.B24 := FALSE;
       #CONTROL_MAN.B25 := FALSE;
       #CONTROL_MAN.B26 := FALSE;
       #CONTROL_MAN.B27 := FALSE;
       #CONTROL_MAN.B28 := FALSE;
       #CONTROL_MAN.B29 := FALSE;
       #CONTROL_MAN.B30 := FALSE;
       #CONTROL_MAN.B31 := FALSE;
       #MEMOR.M6 := TRUE;
       #TRIG.inicial_ok_op := FALSE;
   END_IF;
   #_w2 := NOT "MANUAL" AND #MEMOR.M10;   // falling edge
   #MEMOR.M10 := "MANUAL";
   IF #_w2 THEN #SQCR := #STEP_1000_KONTROLA; END_IF;
   #_w3 := "INICIALIZACE_RUN" AND NOT #MEMOR.M4;   // rising edge
   #MEMOR.M4 := "INICIALIZACE_RUN";
   IF #_w3 THEN #SQCR := #STEP_1000_KONTROLA; END_IF;
END_REGION

REGION Network 3: alarmy
   RUNG wire#powerrail
      { S7_Templates := "SrcType := Int" } NE_Contact(in1 := 0, in2 := "DB_ALARM".OP1."-Y9_ZARAZKA")
      Coil( #MEMOR.M7 )
   END_RUNG
   // the same network as SCL:
   #MEMOR.M7 := 0 <> "DB_ALARM".OP1."-Y9_ZARAZKA";
END_REGION

REGION Network 4: senzory
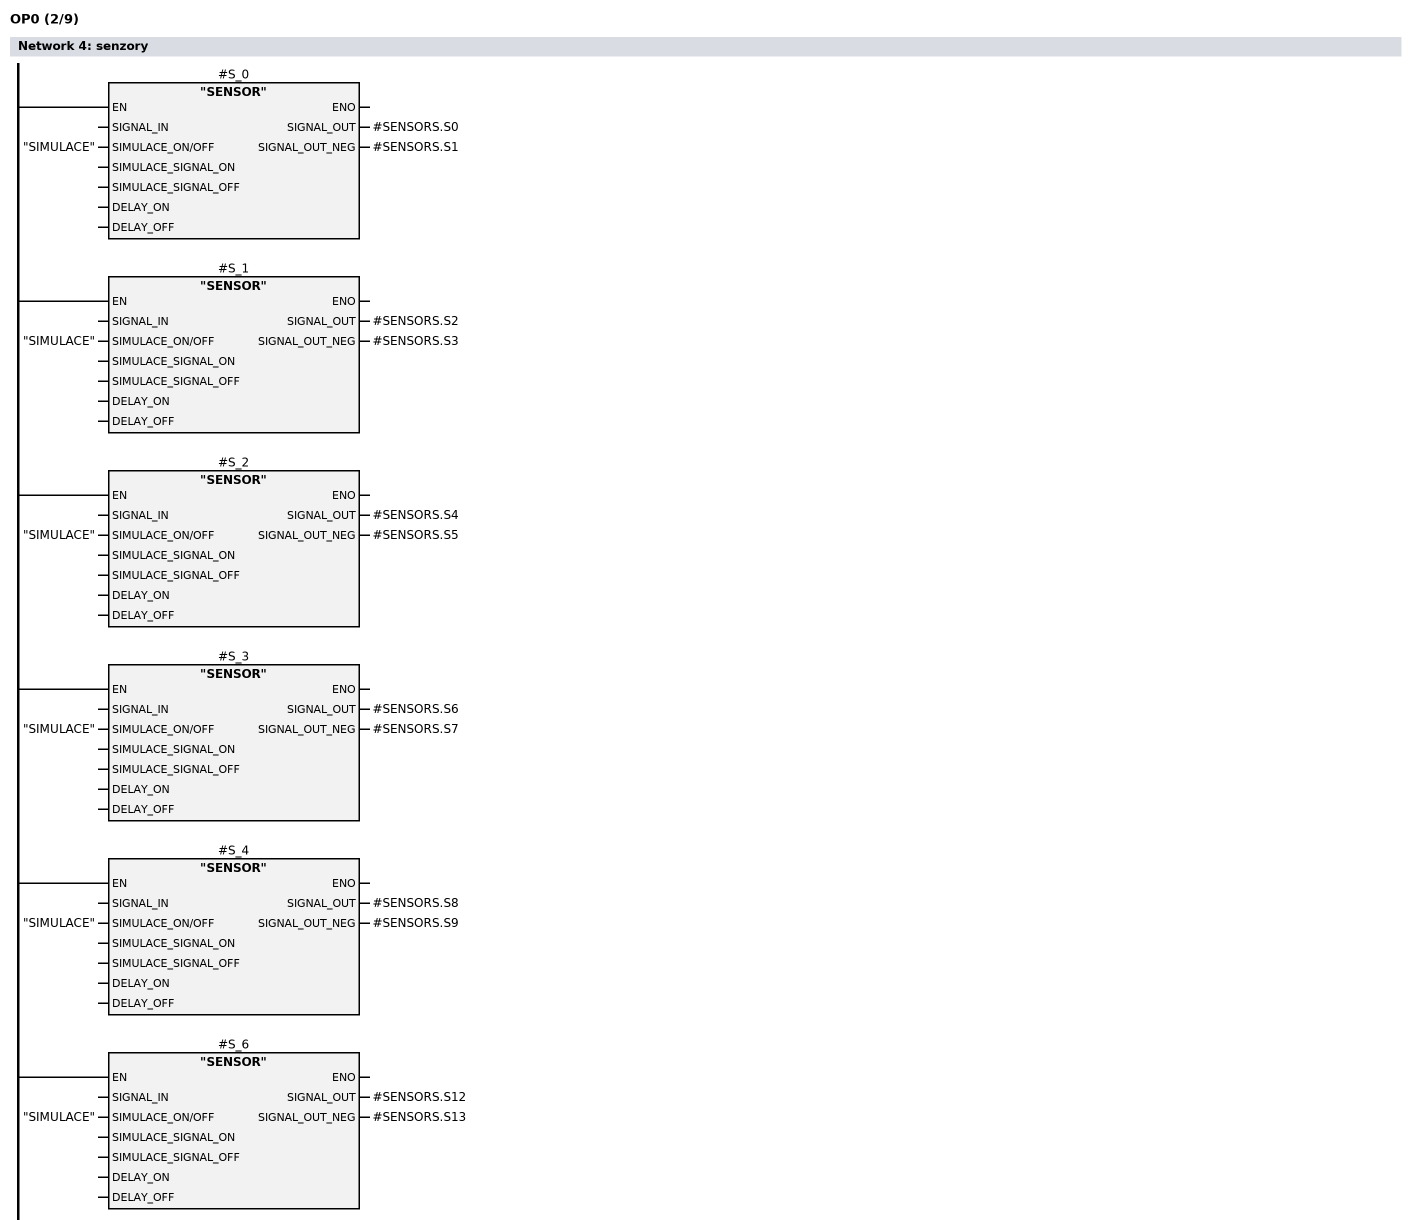
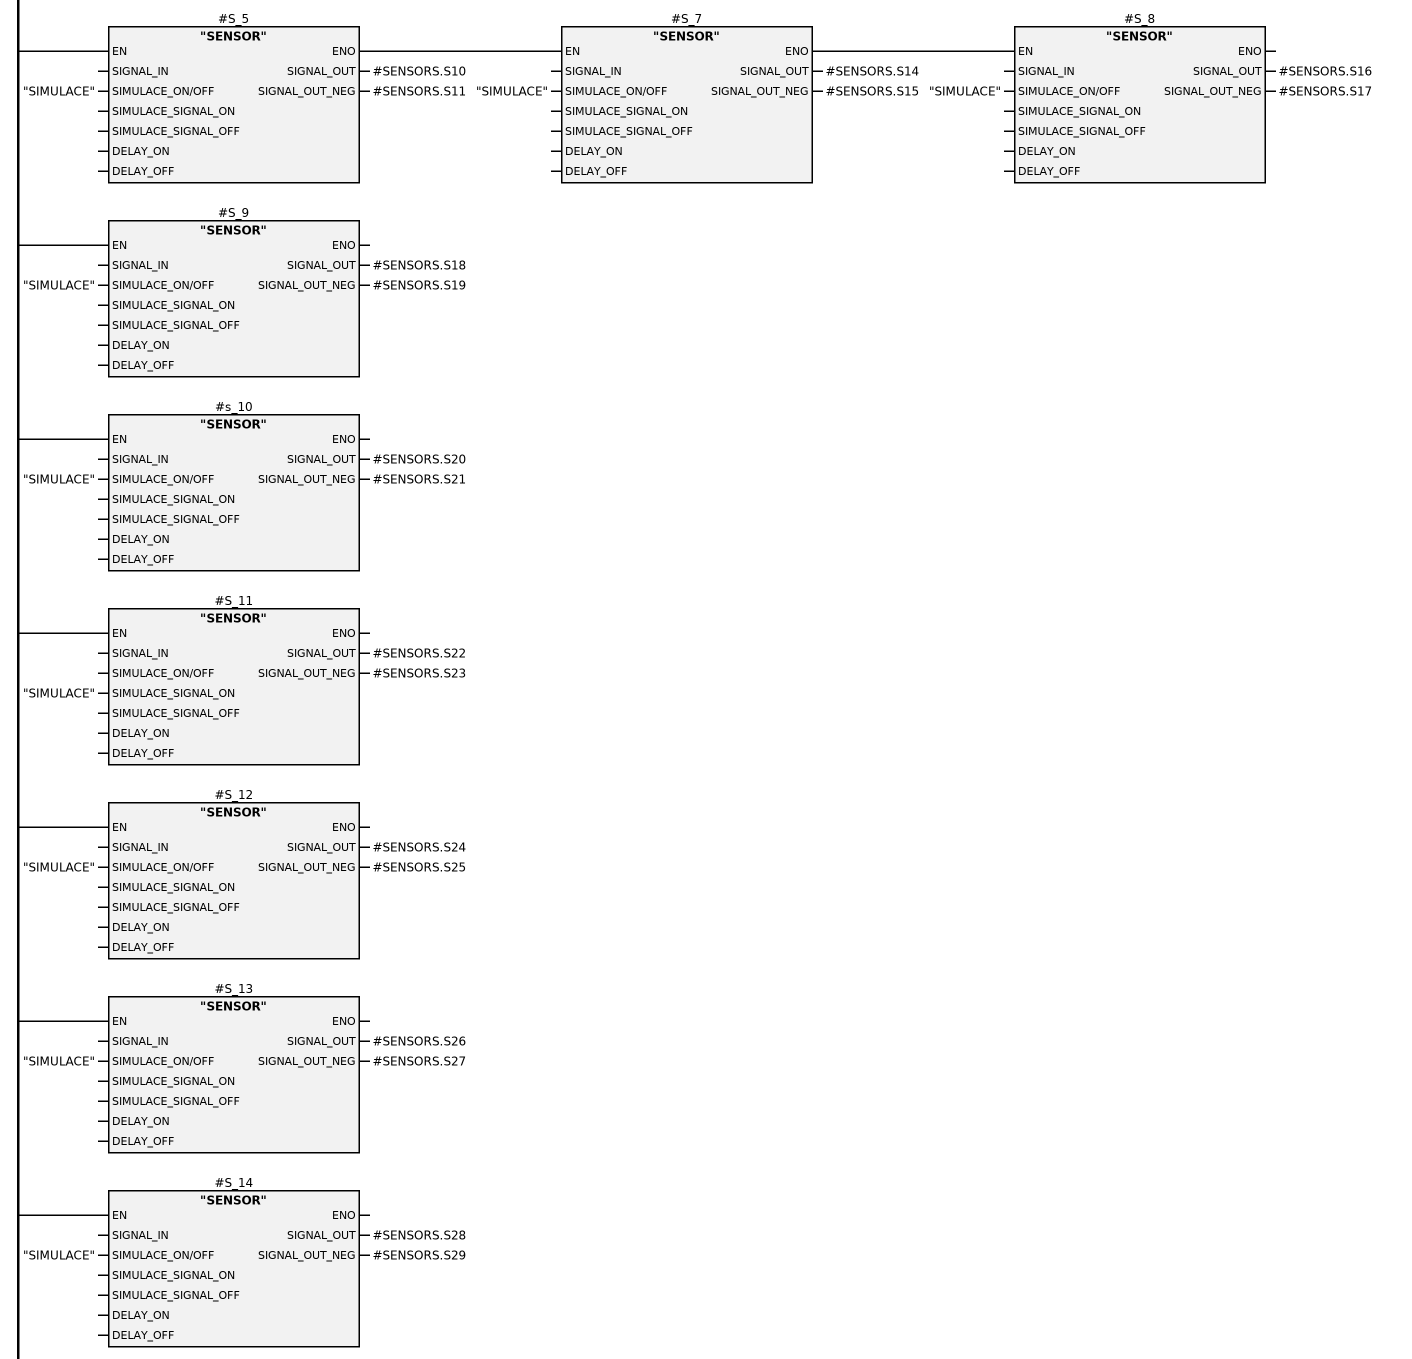
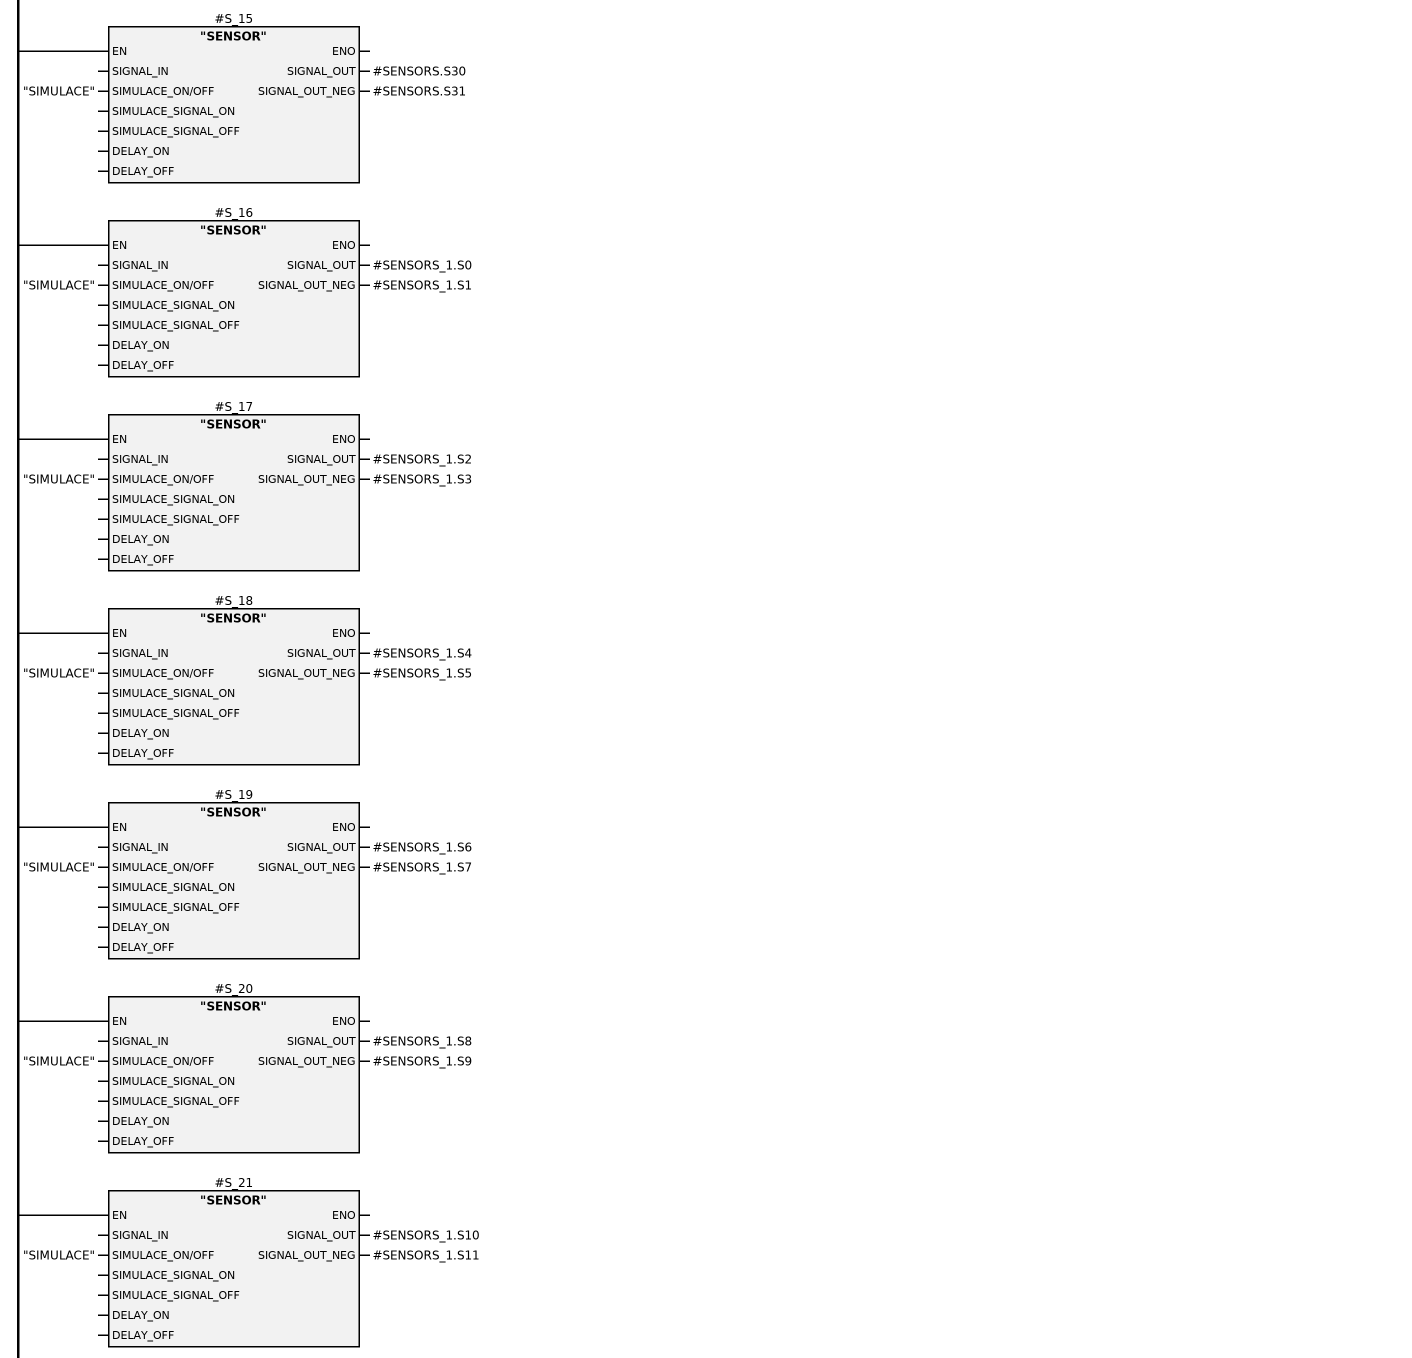
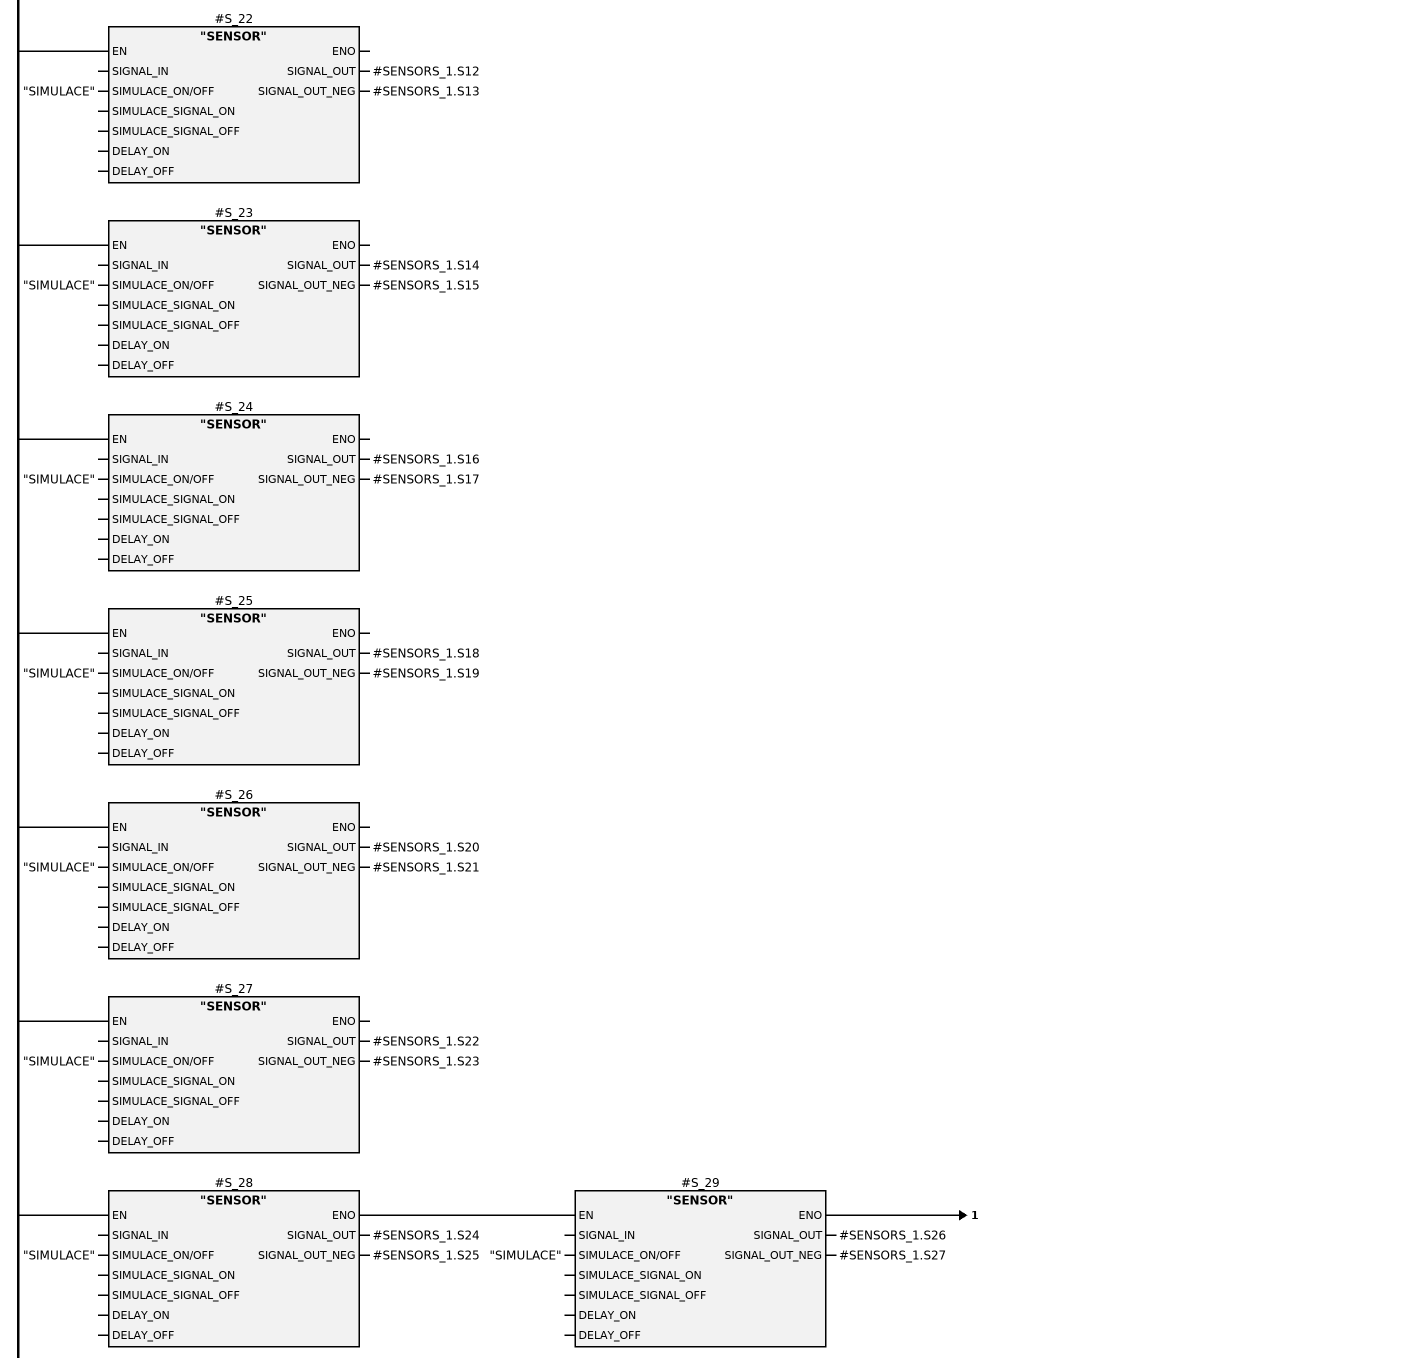
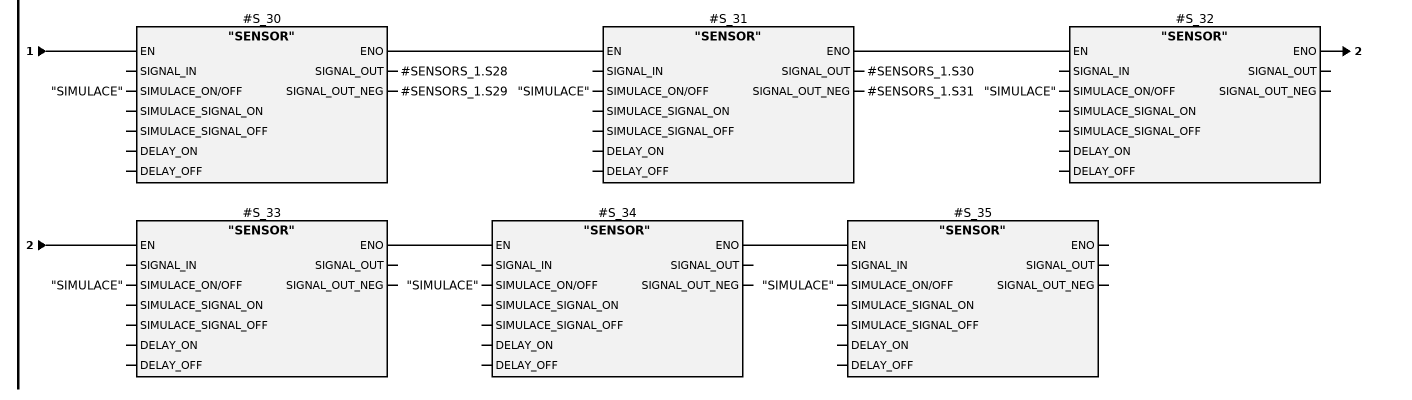
   RUNG wire#powerrail
      #S_0(SIGNAL_IN :=, "SIMULACE_ON/OFF" := "SIMULACE", SIMULACE_SIGNAL_ON :=, SIMULACE_SIGNAL_OFF :=, DELAY_ON :=, DELAY_OFF :=, SIGNAL_OUT => #SENSORS.S0, SIGNAL_OUT_NEG => #SENSORS.S1)
   END_RUNG
   RUNG wire#powerrail
      #S_1(SIGNAL_IN :=, "SIMULACE_ON/OFF" := "SIMULACE", SIMULACE_SIGNAL_ON :=, SIMULACE_SIGNAL_OFF :=, DELAY_ON :=, DELAY_OFF :=, SIGNAL_OUT => #SENSORS.S2, SIGNAL_OUT_NEG => #SENSORS.S3)
   END_RUNG
   RUNG wire#powerrail
      #S_2(SIGNAL_IN :=, "SIMULACE_ON/OFF" := "SIMULACE", SIMULACE_SIGNAL_ON :=, SIMULACE_SIGNAL_OFF :=, DELAY_ON :=, DELAY_OFF :=, SIGNAL_OUT => #SENSORS.S4, SIGNAL_OUT_NEG => #SENSORS.S5)
   END_RUNG
   RUNG wire#powerrail
      #S_3(SIGNAL_IN :=, "SIMULACE_ON/OFF" := "SIMULACE", SIMULACE_SIGNAL_ON :=, SIMULACE_SIGNAL_OFF :=, DELAY_ON :=, DELAY_OFF :=, SIGNAL_OUT => #SENSORS.S6, SIGNAL_OUT_NEG => #SENSORS.S7)
   END_RUNG
   RUNG wire#powerrail
      #S_4(SIGNAL_IN :=, "SIMULACE_ON/OFF" := "SIMULACE", SIMULACE_SIGNAL_ON :=, SIMULACE_SIGNAL_OFF :=, DELAY_ON :=, DELAY_OFF :=, SIGNAL_OUT => #SENSORS.S8, SIGNAL_OUT_NEG => #SENSORS.S9)
   END_RUNG
   RUNG wire#powerrail
      #S_6(SIGNAL_IN :=, "SIMULACE_ON/OFF" := "SIMULACE", SIMULACE_SIGNAL_ON :=, SIMULACE_SIGNAL_OFF :=, DELAY_ON :=, DELAY_OFF :=, SIGNAL_OUT => #SENSORS.S12, SIGNAL_OUT_NEG => #SENSORS.S13)
   END_RUNG
   RUNG wire#powerrail
      #S_5(SIGNAL_IN :=, "SIMULACE_ON/OFF" := "SIMULACE", SIMULACE_SIGNAL_ON :=, SIMULACE_SIGNAL_OFF :=, DELAY_ON :=, DELAY_OFF :=, SIGNAL_OUT => #SENSORS.S10, SIGNAL_OUT_NEG => #SENSORS.S11)
      #S_7(SIGNAL_IN :=, "SIMULACE_ON/OFF" := "SIMULACE", SIMULACE_SIGNAL_ON :=, SIMULACE_SIGNAL_OFF :=, DELAY_ON :=, DELAY_OFF :=, SIGNAL_OUT => #SENSORS.S14, SIGNAL_OUT_NEG => #SENSORS.S15)
      #S_8(SIGNAL_IN :=, "SIMULACE_ON/OFF" := "SIMULACE", SIMULACE_SIGNAL_ON :=, SIMULACE_SIGNAL_OFF :=, DELAY_ON :=, DELAY_OFF :=, SIGNAL_OUT => #SENSORS.S16, SIGNAL_OUT_NEG => #SENSORS.S17)
   END_RUNG
   RUNG wire#powerrail
      #S_9(SIGNAL_IN :=, "SIMULACE_ON/OFF" := "SIMULACE", SIMULACE_SIGNAL_ON :=, SIMULACE_SIGNAL_OFF :=, DELAY_ON :=, DELAY_OFF :=, SIGNAL_OUT => #SENSORS.S18, SIGNAL_OUT_NEG => #SENSORS.S19)
   END_RUNG
   RUNG wire#powerrail
      #s_10(SIGNAL_IN :=, "SIMULACE_ON/OFF" := "SIMULACE", SIMULACE_SIGNAL_ON :=, SIMULACE_SIGNAL_OFF :=, DELAY_ON :=, DELAY_OFF :=, SIGNAL_OUT => #SENSORS.S20, SIGNAL_OUT_NEG => #SENSORS.S21)
   END_RUNG
   RUNG wire#powerrail
      #S_11(SIGNAL_IN :=, "SIMULACE_ON/OFF" :=, SIMULACE_SIGNAL_ON := "SIMULACE", SIMULACE_SIGNAL_OFF :=, DELAY_ON :=, DELAY_OFF :=, SIGNAL_OUT => #SENSORS.S22, SIGNAL_OUT_NEG => #SENSORS.S23)
   END_RUNG
   RUNG wire#powerrail
      #S_12(SIGNAL_IN :=, "SIMULACE_ON/OFF" := "SIMULACE", SIMULACE_SIGNAL_ON :=, SIMULACE_SIGNAL_OFF :=, DELAY_ON :=, DELAY_OFF :=, SIGNAL_OUT => #SENSORS.S24, SIGNAL_OUT_NEG => #SENSORS.S25)
   END_RUNG
   RUNG wire#powerrail
      #S_13(SIGNAL_IN :=, "SIMULACE_ON/OFF" := "SIMULACE", SIMULACE_SIGNAL_ON :=, SIMULACE_SIGNAL_OFF :=, DELAY_ON :=, DELAY_OFF :=, SIGNAL_OUT => #SENSORS.S26, SIGNAL_OUT_NEG => #SENSORS.S27)
   END_RUNG
   RUNG wire#powerrail
      #S_14(SIGNAL_IN :=, "SIMULACE_ON/OFF" := "SIMULACE", SIMULACE_SIGNAL_ON :=, SIMULACE_SIGNAL_OFF :=, DELAY_ON :=, DELAY_OFF :=, SIGNAL_OUT => #SENSORS.S28, SIGNAL_OUT_NEG => #SENSORS.S29)
   END_RUNG
   RUNG wire#powerrail
      #S_15(SIGNAL_IN :=, "SIMULACE_ON/OFF" := "SIMULACE", SIMULACE_SIGNAL_ON :=, SIMULACE_SIGNAL_OFF :=, DELAY_ON :=, DELAY_OFF :=, SIGNAL_OUT => #SENSORS.S30, SIGNAL_OUT_NEG => #SENSORS.S31)
   END_RUNG
   RUNG wire#powerrail
      #S_16(SIGNAL_IN :=, "SIMULACE_ON/OFF" := "SIMULACE", SIMULACE_SIGNAL_ON :=, SIMULACE_SIGNAL_OFF :=, DELAY_ON :=, DELAY_OFF :=, SIGNAL_OUT => #SENSORS_1.S0, SIGNAL_OUT_NEG => #SENSORS_1.S1)
   END_RUNG
   RUNG wire#powerrail
      #S_17(SIGNAL_IN :=, "SIMULACE_ON/OFF" := "SIMULACE", SIMULACE_SIGNAL_ON :=, SIMULACE_SIGNAL_OFF :=, DELAY_ON :=, DELAY_OFF :=, SIGNAL_OUT => #SENSORS_1.S2, SIGNAL_OUT_NEG => #SENSORS_1.S3)
   END_RUNG
   RUNG wire#powerrail
      #S_18(SIGNAL_IN :=, "SIMULACE_ON/OFF" := "SIMULACE", SIMULACE_SIGNAL_ON :=, SIMULACE_SIGNAL_OFF :=, DELAY_ON :=, DELAY_OFF :=, SIGNAL_OUT => #SENSORS_1.S4, SIGNAL_OUT_NEG => #SENSORS_1.S5)
   END_RUNG
   RUNG wire#powerrail
      #S_19(SIGNAL_IN :=, "SIMULACE_ON/OFF" := "SIMULACE", SIMULACE_SIGNAL_ON :=, SIMULACE_SIGNAL_OFF :=, DELAY_ON :=, DELAY_OFF :=, SIGNAL_OUT => #SENSORS_1.S6, SIGNAL_OUT_NEG => #SENSORS_1.S7)
   END_RUNG
   RUNG wire#powerrail
      #S_20(SIGNAL_IN :=, "SIMULACE_ON/OFF" := "SIMULACE", SIMULACE_SIGNAL_ON :=, SIMULACE_SIGNAL_OFF :=, DELAY_ON :=, DELAY_OFF :=, SIGNAL_OUT => #SENSORS_1.S8, SIGNAL_OUT_NEG => #SENSORS_1.S9)
   END_RUNG
   RUNG wire#powerrail
      #S_21(SIGNAL_IN :=, "SIMULACE_ON/OFF" := "SIMULACE", SIMULACE_SIGNAL_ON :=, SIMULACE_SIGNAL_OFF :=, DELAY_ON :=, DELAY_OFF :=, SIGNAL_OUT => #SENSORS_1.S10, SIGNAL_OUT_NEG => #SENSORS_1.S11)
   END_RUNG
   RUNG wire#powerrail
      #S_22(SIGNAL_IN :=, "SIMULACE_ON/OFF" := "SIMULACE", SIMULACE_SIGNAL_ON :=, SIMULACE_SIGNAL_OFF :=, DELAY_ON :=, DELAY_OFF :=, SIGNAL_OUT => #SENSORS_1.S12, SIGNAL_OUT_NEG => #SENSORS_1.S13)
   END_RUNG
   RUNG wire#powerrail
      #S_23(SIGNAL_IN :=, "SIMULACE_ON/OFF" := "SIMULACE", SIMULACE_SIGNAL_ON :=, SIMULACE_SIGNAL_OFF :=, DELAY_ON :=, DELAY_OFF :=, SIGNAL_OUT => #SENSORS_1.S14, SIGNAL_OUT_NEG => #SENSORS_1.S15)
   END_RUNG
   RUNG wire#powerrail
      #S_24(SIGNAL_IN :=, "SIMULACE_ON/OFF" := "SIMULACE", SIMULACE_SIGNAL_ON :=, SIMULACE_SIGNAL_OFF :=, DELAY_ON :=, DELAY_OFF :=, SIGNAL_OUT => #SENSORS_1.S16, SIGNAL_OUT_NEG => #SENSORS_1.S17)
   END_RUNG
   RUNG wire#powerrail
      #S_25(SIGNAL_IN :=, "SIMULACE_ON/OFF" := "SIMULACE", SIMULACE_SIGNAL_ON :=, SIMULACE_SIGNAL_OFF :=, DELAY_ON :=, DELAY_OFF :=, SIGNAL_OUT => #SENSORS_1.S18, SIGNAL_OUT_NEG => #SENSORS_1.S19)
   END_RUNG
   RUNG wire#powerrail
      #S_26(SIGNAL_IN :=, "SIMULACE_ON/OFF" := "SIMULACE", SIMULACE_SIGNAL_ON :=, SIMULACE_SIGNAL_OFF :=, DELAY_ON :=, DELAY_OFF :=, SIGNAL_OUT => #SENSORS_1.S20, SIGNAL_OUT_NEG => #SENSORS_1.S21)
   END_RUNG
   RUNG wire#powerrail
      #S_27(SIGNAL_IN :=, "SIMULACE_ON/OFF" := "SIMULACE", SIMULACE_SIGNAL_ON :=, SIMULACE_SIGNAL_OFF :=, DELAY_ON :=, DELAY_OFF :=, SIGNAL_OUT => #SENSORS_1.S22, SIGNAL_OUT_NEG => #SENSORS_1.S23)
   END_RUNG
   RUNG wire#powerrail
      #S_28(SIGNAL_IN :=, "SIMULACE_ON/OFF" := "SIMULACE", SIMULACE_SIGNAL_ON :=, SIMULACE_SIGNAL_OFF :=, DELAY_ON :=, DELAY_OFF :=, SIGNAL_OUT => #SENSORS_1.S24, SIGNAL_OUT_NEG => #SENSORS_1.S25)
      #S_29(SIGNAL_IN :=, "SIMULACE_ON/OFF" := "SIMULACE", SIMULACE_SIGNAL_ON :=, SIMULACE_SIGNAL_OFF :=, DELAY_ON :=, DELAY_OFF :=, SIGNAL_OUT => #SENSORS_1.S26, SIGNAL_OUT_NEG => #SENSORS_1.S27)
      #S_30(SIGNAL_IN :=, "SIMULACE_ON/OFF" := "SIMULACE", SIMULACE_SIGNAL_ON :=, SIMULACE_SIGNAL_OFF :=, DELAY_ON :=, DELAY_OFF :=, SIGNAL_OUT => #SENSORS_1.S28, SIGNAL_OUT_NEG => #SENSORS_1.S29)
      #S_31(SIGNAL_IN :=, "SIMULACE_ON/OFF" := "SIMULACE", SIMULACE_SIGNAL_ON :=, SIMULACE_SIGNAL_OFF :=, DELAY_ON :=, DELAY_OFF :=, SIGNAL_OUT => #SENSORS_1.S30, SIGNAL_OUT_NEG => #SENSORS_1.S31)
      #S_32(SIGNAL_IN :=, "SIMULACE_ON/OFF" := "SIMULACE", SIMULACE_SIGNAL_ON :=, SIMULACE_SIGNAL_OFF :=, DELAY_ON :=, DELAY_OFF :=, SIGNAL_OUT =>, SIGNAL_OUT_NEG =>)
      #S_33(SIGNAL_IN :=, "SIMULACE_ON/OFF" := "SIMULACE", SIMULACE_SIGNAL_ON :=, SIMULACE_SIGNAL_OFF :=, DELAY_ON :=, DELAY_OFF :=, SIGNAL_OUT =>, SIGNAL_OUT_NEG =>)
      #S_34(SIGNAL_IN :=, "SIMULACE_ON/OFF" := "SIMULACE", SIMULACE_SIGNAL_ON :=, SIMULACE_SIGNAL_OFF :=, DELAY_ON :=, DELAY_OFF :=, SIGNAL_OUT =>, SIGNAL_OUT_NEG =>)
      #S_35(SIGNAL_IN :=, "SIMULACE_ON/OFF" := "SIMULACE", SIMULACE_SIGNAL_ON :=, SIMULACE_SIGNAL_OFF :=, DELAY_ON :=, DELAY_OFF :=, SIGNAL_OUT =>, SIGNAL_OUT_NEG =>)
   END_RUNG
   // the same network as SCL:
   #S_0("SIMULACE_ON/OFF" := "SIMULACE", SIGNAL_OUT => #SENSORS.S0, SIGNAL_OUT_NEG => #SENSORS.S1);   // "SENSOR"
   #S_1("SIMULACE_ON/OFF" := "SIMULACE", SIGNAL_OUT => #SENSORS.S2, SIGNAL_OUT_NEG => #SENSORS.S3);   // "SENSOR"
   #S_2("SIMULACE_ON/OFF" := "SIMULACE", SIGNAL_OUT => #SENSORS.S4, SIGNAL_OUT_NEG => #SENSORS.S5);   // "SENSOR"
   #S_3("SIMULACE_ON/OFF" := "SIMULACE", SIGNAL_OUT => #SENSORS.S6, SIGNAL_OUT_NEG => #SENSORS.S7);   // "SENSOR"
   #S_4("SIMULACE_ON/OFF" := "SIMULACE", SIGNAL_OUT => #SENSORS.S8, SIGNAL_OUT_NEG => #SENSORS.S9);   // "SENSOR"
   #S_6("SIMULACE_ON/OFF" := "SIMULACE", SIGNAL_OUT => #SENSORS.S12, SIGNAL_OUT_NEG => #SENSORS.S13);   // "SENSOR"
   #S_5("SIMULACE_ON/OFF" := "SIMULACE",   // "SENSOR"
        SIGNAL_OUT => #SENSORS.S10,
        SIGNAL_OUT_NEG => #SENSORS.S11,
        ENO => #_w1);
   #S_7(EN := #_w1,   // "SENSOR"
        "SIMULACE_ON/OFF" := "SIMULACE",
        SIGNAL_OUT => #SENSORS.S14,
        SIGNAL_OUT_NEG => #SENSORS.S15,
        ENO => #_w2);
   IF #_w2 THEN
       #S_8("SIMULACE_ON/OFF" := "SIMULACE", SIGNAL_OUT => #SENSORS.S16, SIGNAL_OUT_NEG => #SENSORS.S17);   // "SENSOR"
   END_IF;
   #S_9("SIMULACE_ON/OFF" := "SIMULACE", SIGNAL_OUT => #SENSORS.S18, SIGNAL_OUT_NEG => #SENSORS.S19);   // "SENSOR"
   #s_10("SIMULACE_ON/OFF" := "SIMULACE", SIGNAL_OUT => #SENSORS.S20, SIGNAL_OUT_NEG => #SENSORS.S21);   // "SENSOR"
   #S_11(SIMULACE_SIGNAL_ON := "SIMULACE", SIGNAL_OUT => #SENSORS.S22, SIGNAL_OUT_NEG => #SENSORS.S23);   // "SENSOR"
   #S_12("SIMULACE_ON/OFF" := "SIMULACE", SIGNAL_OUT => #SENSORS.S24, SIGNAL_OUT_NEG => #SENSORS.S25);   // "SENSOR"
   #S_13("SIMULACE_ON/OFF" := "SIMULACE", SIGNAL_OUT => #SENSORS.S26, SIGNAL_OUT_NEG => #SENSORS.S27);   // "SENSOR"
   #S_14("SIMULACE_ON/OFF" := "SIMULACE", SIGNAL_OUT => #SENSORS.S28, SIGNAL_OUT_NEG => #SENSORS.S29);   // "SENSOR"
   #S_15("SIMULACE_ON/OFF" := "SIMULACE", SIGNAL_OUT => #SENSORS.S30, SIGNAL_OUT_NEG => #SENSORS.S31);   // "SENSOR"
   #S_16("SIMULACE_ON/OFF" := "SIMULACE", SIGNAL_OUT => #SENSORS_1.S0, SIGNAL_OUT_NEG => #SENSORS_1.S1);   // "SENSOR"
   #S_17("SIMULACE_ON/OFF" := "SIMULACE", SIGNAL_OUT => #SENSORS_1.S2, SIGNAL_OUT_NEG => #SENSORS_1.S3);   // "SENSOR"
   #S_18("SIMULACE_ON/OFF" := "SIMULACE", SIGNAL_OUT => #SENSORS_1.S4, SIGNAL_OUT_NEG => #SENSORS_1.S5);   // "SENSOR"
   #S_19("SIMULACE_ON/OFF" := "SIMULACE", SIGNAL_OUT => #SENSORS_1.S6, SIGNAL_OUT_NEG => #SENSORS_1.S7);   // "SENSOR"
   #S_20("SIMULACE_ON/OFF" := "SIMULACE", SIGNAL_OUT => #SENSORS_1.S8, SIGNAL_OUT_NEG => #SENSORS_1.S9);   // "SENSOR"
   #S_21("SIMULACE_ON/OFF" := "SIMULACE", SIGNAL_OUT => #SENSORS_1.S10, SIGNAL_OUT_NEG => #SENSORS_1.S11);   // "SENSOR"
   #S_22("SIMULACE_ON/OFF" := "SIMULACE", SIGNAL_OUT => #SENSORS_1.S12, SIGNAL_OUT_NEG => #SENSORS_1.S13);   // "SENSOR"
   #S_23("SIMULACE_ON/OFF" := "SIMULACE", SIGNAL_OUT => #SENSORS_1.S14, SIGNAL_OUT_NEG => #SENSORS_1.S15);   // "SENSOR"
   #S_24("SIMULACE_ON/OFF" := "SIMULACE", SIGNAL_OUT => #SENSORS_1.S16, SIGNAL_OUT_NEG => #SENSORS_1.S17);   // "SENSOR"
   #S_25("SIMULACE_ON/OFF" := "SIMULACE", SIGNAL_OUT => #SENSORS_1.S18, SIGNAL_OUT_NEG => #SENSORS_1.S19);   // "SENSOR"
   #S_26("SIMULACE_ON/OFF" := "SIMULACE", SIGNAL_OUT => #SENSORS_1.S20, SIGNAL_OUT_NEG => #SENSORS_1.S21);   // "SENSOR"
   #S_27("SIMULACE_ON/OFF" := "SIMULACE", SIGNAL_OUT => #SENSORS_1.S22, SIGNAL_OUT_NEG => #SENSORS_1.S23);   // "SENSOR"
   #S_28("SIMULACE_ON/OFF" := "SIMULACE",   // "SENSOR"
         SIGNAL_OUT => #SENSORS_1.S24,
         SIGNAL_OUT_NEG => #SENSORS_1.S25,
         ENO => #_w3);
   #S_29(EN := #_w3,   // "SENSOR"
         "SIMULACE_ON/OFF" := "SIMULACE",
         SIGNAL_OUT => #SENSORS_1.S26,
         SIGNAL_OUT_NEG => #SENSORS_1.S27,
         ENO => #_w4);
   #S_30(EN := #_w4,   // "SENSOR"
         "SIMULACE_ON/OFF" := "SIMULACE",
         SIGNAL_OUT => #SENSORS_1.S28,
         SIGNAL_OUT_NEG => #SENSORS_1.S29,
         ENO => #_w5);
   #S_31(EN := #_w5,   // "SENSOR"
         "SIMULACE_ON/OFF" := "SIMULACE",
         SIGNAL_OUT => #SENSORS_1.S30,
         SIGNAL_OUT_NEG => #SENSORS_1.S31,
         ENO => #_w6);
   #S_32(EN := #_w6, "SIMULACE_ON/OFF" := "SIMULACE", ENO => #_w7);   // "SENSOR"
   #S_33(EN := #_w7, "SIMULACE_ON/OFF" := "SIMULACE", ENO => #_w8);   // "SENSOR"
   #S_34(EN := #_w8, "SIMULACE_ON/OFF" := "SIMULACE", ENO => #_w9);   // "SENSOR"
   IF #_w9 THEN
       #S_35("SIMULACE_ON/OFF" := "SIMULACE");   // "SENSOR"
   END_IF;
END_REGION

REGION Network 5: INICIALIZACE START
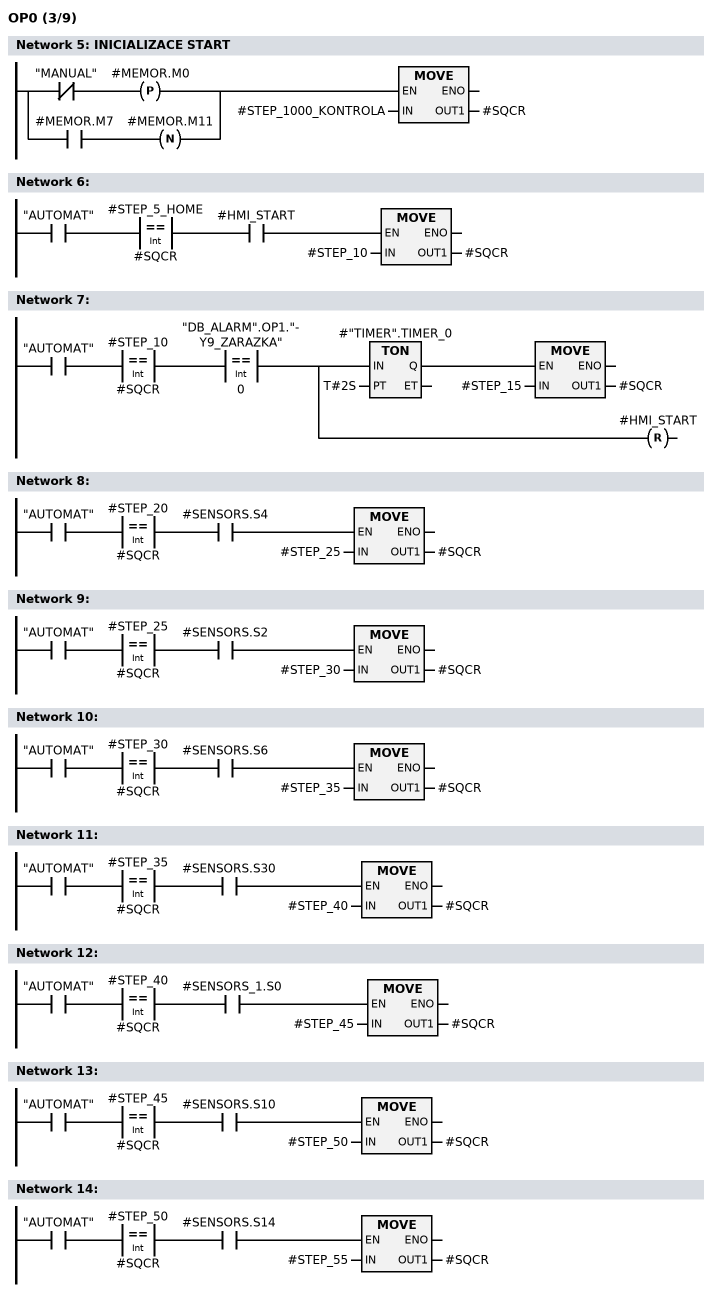
   RUNG wire#powerrail
      I_Contact( "MANUAL" )
      P_Trig( #MEMOR.M0 )
      wire#w1
      Move(in := #STEP_1000_KONTROLA, out1 => #SQCR)
   END_RUNG
   RUNG wire#powerrail
      Contact( #MEMOR.M7 )
      N_Trig( #MEMOR.M11 )
   END_RUNG wire#w1
   // the same network as SCL:
   #_w1 := NOT "MANUAL" AND NOT #MEMOR.M0;   // rising edge
   #MEMOR.M0 := NOT "MANUAL";
   #_w2 := NOT #MEMOR.M7 AND #MEMOR.M11;   // falling edge
   #MEMOR.M11 := #MEMOR.M7;
   IF #_w1 OR #_w2 THEN #SQCR := #STEP_1000_KONTROLA; END_IF;
END_REGION

REGION Network 6
   RUNG wire#powerrail
      Contact( "AUTOMAT" )
      { S7_Templates := "SrcType := Int" } EQ_Contact(in1 := #STEP_5_HOME, in2 := #SQCR)
      Contact( #HMI_START )
      Move(in := #STEP_10, out1 => #SQCR)
   END_RUNG
   // the same network as SCL:
   IF "AUTOMAT" AND (#STEP_5_HOME = #SQCR) AND #HMI_START THEN #SQCR := #STEP_10; END_IF;
END_REGION

REGION Network 7
   #_w1 := "AUTOMAT" AND (#STEP_10 = #SQCR) AND ("DB_ALARM".OP1."-Y9_ZARAZKA" = 0);
   #"TIMER".TIMER_0.TON(IN := #_w1, PT := T#2S);
   IF #"TIMER".TIMER_0.Q THEN #SQCR := #STEP_15; END_IF;
   IF #_w1 THEN #HMI_START := FALSE; END_IF;
END_REGION

REGION Network 8
   RUNG wire#powerrail
      Contact( "AUTOMAT" )
      { S7_Templates := "SrcType := Int" } EQ_Contact(in1 := #STEP_20, in2 := #SQCR)
      Contact( #SENSORS.S4 )
      Move(in := #STEP_25, out1 => #SQCR)
   END_RUNG
   // the same network as SCL:
   IF "AUTOMAT" AND (#STEP_20 = #SQCR) AND #SENSORS.S4 THEN #SQCR := #STEP_25; END_IF;
END_REGION

REGION Network 9
   RUNG wire#powerrail
      Contact( "AUTOMAT" )
      { S7_Templates := "SrcType := Int" } EQ_Contact(in1 := #STEP_25, in2 := #SQCR)
      Contact( #SENSORS.S2 )
      Move(in := #STEP_30, out1 => #SQCR)
   END_RUNG
   // the same network as SCL:
   IF "AUTOMAT" AND (#STEP_25 = #SQCR) AND #SENSORS.S2 THEN #SQCR := #STEP_30; END_IF;
END_REGION

REGION Network 10
   RUNG wire#powerrail
      Contact( "AUTOMAT" )
      { S7_Templates := "SrcType := Int" } EQ_Contact(in1 := #STEP_30, in2 := #SQCR)
      Contact( #SENSORS.S6 )
      Move(in := #STEP_35, out1 => #SQCR)
   END_RUNG
   // the same network as SCL:
   IF "AUTOMAT" AND (#STEP_30 = #SQCR) AND #SENSORS.S6 THEN #SQCR := #STEP_35; END_IF;
END_REGION

REGION Network 11
   RUNG wire#powerrail
      Contact( "AUTOMAT" )
      { S7_Templates := "SrcType := Int" } EQ_Contact(in1 := #STEP_35, in2 := #SQCR)
      Contact( #SENSORS.S30 )
      Move(in := #STEP_40, out1 => #SQCR)
   END_RUNG
   // the same network as SCL:
   IF "AUTOMAT" AND (#STEP_35 = #SQCR) AND #SENSORS.S30 THEN #SQCR := #STEP_40; END_IF;
END_REGION

REGION Network 12
   RUNG wire#powerrail
      Contact( "AUTOMAT" )
      { S7_Templates := "SrcType := Int" } EQ_Contact(in1 := #STEP_40, in2 := #SQCR)
      Contact( #SENSORS_1.S0 )
      Move(in := #STEP_45, out1 => #SQCR)
   END_RUNG
   // the same network as SCL:
   IF "AUTOMAT" AND (#STEP_40 = #SQCR) AND #SENSORS_1.S0 THEN #SQCR := #STEP_45; END_IF;
END_REGION

REGION Network 13
   RUNG wire#powerrail
      Contact( "AUTOMAT" )
      { S7_Templates := "SrcType := Int" } EQ_Contact(in1 := #STEP_45, in2 := #SQCR)
      Contact( #SENSORS.S10 )
      Move(in := #STEP_50, out1 => #SQCR)
   END_RUNG
   // the same network as SCL:
   IF "AUTOMAT" AND (#STEP_45 = #SQCR) AND #SENSORS.S10 THEN #SQCR := #STEP_50; END_IF;
END_REGION

REGION Network 14
   RUNG wire#powerrail
      Contact( "AUTOMAT" )
      { S7_Templates := "SrcType := Int" } EQ_Contact(in1 := #STEP_50, in2 := #SQCR)
      Contact( #SENSORS.S14 )
      Move(in := #STEP_55, out1 => #SQCR)
   END_RUNG
   // the same network as SCL:
   IF "AUTOMAT" AND (#STEP_50 = #SQCR) AND #SENSORS.S14 THEN #SQCR := #STEP_55; END_IF;
END_REGION

REGION Network 15
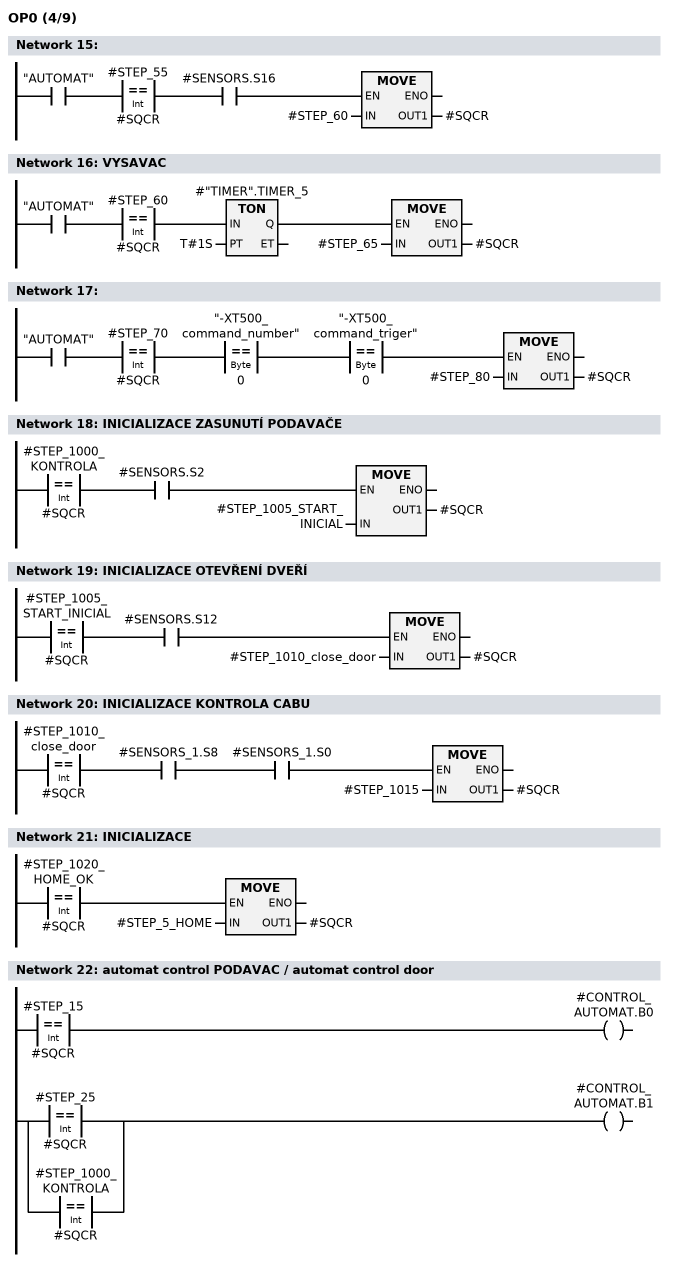
   RUNG wire#powerrail
      Contact( "AUTOMAT" )
      { S7_Templates := "SrcType := Int" } EQ_Contact(in1 := #STEP_55, in2 := #SQCR)
      Contact( #SENSORS.S16 )
      Move(in := #STEP_60, out1 => #SQCR)
   END_RUNG
   // the same network as SCL:
   IF "AUTOMAT" AND (#STEP_55 = #SQCR) AND #SENSORS.S16 THEN #SQCR := #STEP_60; END_IF;
END_REGION

REGION Network 16: VYSAVAC
   #"TIMER".TIMER_5.TON(IN := "AUTOMAT" AND (#STEP_60 = #SQCR), PT := T#1S);
   IF #"TIMER".TIMER_5.Q THEN #SQCR := #STEP_65; END_IF;
END_REGION

REGION Network 17
   RUNG wire#powerrail
      Contact( "AUTOMAT" )
      { S7_Templates := "SrcType := Int" } EQ_Contact(in1 := #STEP_70, in2 := #SQCR)
      { S7_Templates := "SrcType := Byte" } EQ_Contact(in1 := "-XT500_command_number", in2 := 0)
      { S7_Templates := "SrcType := Byte" } EQ_Contact(in1 := "-XT500_command_triger", in2 := 0)
      Move(in := #STEP_80, out1 => #SQCR)
   END_RUNG
   // the same network as SCL:
   IF "AUTOMAT" AND (#STEP_70 = #SQCR) AND ("-XT500_command_number" = 0) AND ("-XT500_command_triger" = 0) THEN
       #SQCR := #STEP_80;
   END_IF;
END_REGION

REGION Network 18: INICIALIZACE ZASUNUTÍ PODAVAČE
   RUNG wire#powerrail
      { S7_Templates := "SrcType := Int" } EQ_Contact(in1 := #STEP_1000_KONTROLA, in2 := #SQCR)
      Contact( #SENSORS.S2 )
      Move(in := #STEP_1005_START_INICIAL, out1 => #SQCR)
   END_RUNG
   // the same network as SCL:
   IF (#STEP_1000_KONTROLA = #SQCR) AND #SENSORS.S2 THEN #SQCR := #STEP_1005_START_INICIAL; END_IF;
END_REGION

REGION Network 19: INICIALIZACE OTEVŘENÍ DVEŘÍ
   RUNG wire#powerrail
      { S7_Templates := "SrcType := Int" } EQ_Contact(in1 := #STEP_1005_START_INICIAL, in2 := #SQCR)
      Contact( #SENSORS.S12 )
      Move(in := #STEP_1010_close_door, out1 => #SQCR)
   END_RUNG
   // the same network as SCL:
   IF (#STEP_1005_START_INICIAL = #SQCR) AND #SENSORS.S12 THEN #SQCR := #STEP_1010_close_door; END_IF;
END_REGION

REGION Network 20: INICIALIZACE KONTROLA CABU
   RUNG wire#powerrail
      { S7_Templates := "SrcType := Int" } EQ_Contact(in1 := #STEP_1010_close_door, in2 := #SQCR)
      Contact( #SENSORS_1.S8 )
      Contact( #SENSORS_1.S0 )
      Move(in := #STEP_1015, out1 => #SQCR)
   END_RUNG
   // the same network as SCL:
   IF (#STEP_1010_close_door = #SQCR) AND #SENSORS_1.S8 AND #SENSORS_1.S0 THEN #SQCR := #STEP_1015; END_IF;
END_REGION

REGION Network 21: INICIALIZACE
   RUNG wire#powerrail
      { S7_Templates := "SrcType := Int" } EQ_Contact(in1 := #STEP_1020_HOME_OK, in2 := #SQCR)
      Move(in := #STEP_5_HOME, out1 => #SQCR)
   END_RUNG
   // the same network as SCL:
   IF #STEP_1020_HOME_OK = #SQCR THEN #SQCR := #STEP_5_HOME; END_IF;
END_REGION

REGION Network 22: automat control PODAVAC / automat control door
   RUNG wire#powerrail
      { S7_Templates := "SrcType := Int" } EQ_Contact(in1 := #STEP_15, in2 := #SQCR)
      Coil( #CONTROL_AUTOMAT.B0 )
   END_RUNG
   RUNG wire#powerrail
      { S7_Templates := "SrcType := Int" } EQ_Contact(in1 := #STEP_25, in2 := #SQCR)
      wire#w1
      Coil( #CONTROL_AUTOMAT.B1 )
   END_RUNG
   RUNG wire#powerrail
      { S7_Templates := "SrcType := Int" } EQ_Contact(in1 := #STEP_1000_KONTROLA, in2 := #SQCR)
   END_RUNG wire#w1
   // the same network as SCL:
   #CONTROL_AUTOMAT.B0 := #STEP_15 = #SQCR;
   #CONTROL_AUTOMAT.B1 := (#STEP_25 = #SQCR) OR (#STEP_1000_KONTROLA = #SQCR);
END_REGION

REGION Network 23: automat controlMOTOR / automat control osa Z
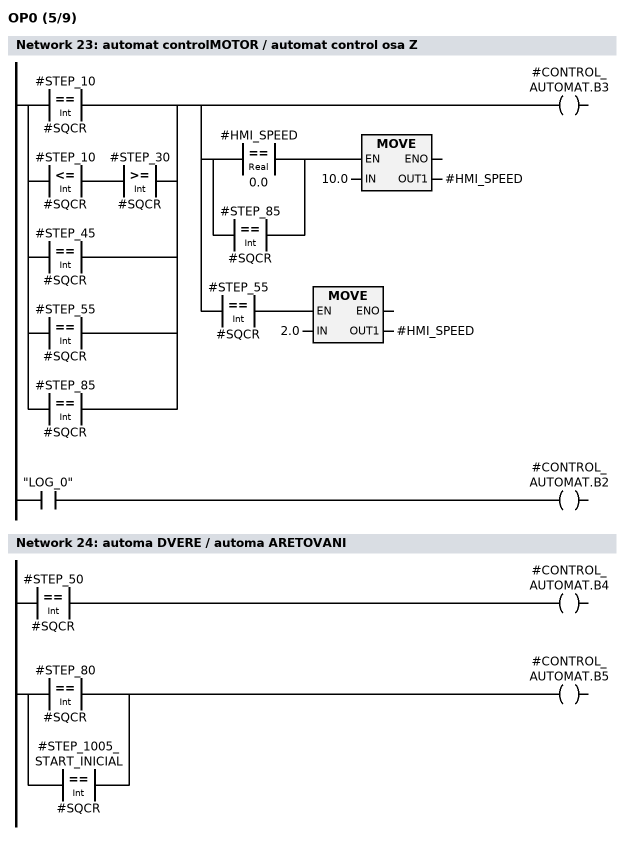
   RUNG wire#powerrail
      { S7_Templates := "SrcType := Int" } EQ_Contact(in1 := #STEP_10, in2 := #SQCR)
      wire#w1
      Coil( #CONTROL_AUTOMAT.B3 )
   END_RUNG
   RUNG wire#powerrail
      { S7_Templates := "SrcType := Int" } LE_Contact(in1 := #STEP_10, in2 := #SQCR)
      { S7_Templates := "SrcType := Int" } GE_Contact(in1 := #STEP_30, in2 := #SQCR)
   END_RUNG wire#w1
   RUNG wire#powerrail
      { S7_Templates := "SrcType := Int" } EQ_Contact(in1 := #STEP_45, in2 := #SQCR)
   END_RUNG wire#w1
   RUNG wire#powerrail
      { S7_Templates := "SrcType := Int" } EQ_Contact(in1 := #STEP_55, in2 := #SQCR)
   END_RUNG wire#w1
   RUNG wire#powerrail
      { S7_Templates := "SrcType := Int" } EQ_Contact(in1 := #STEP_85, in2 := #SQCR)
   END_RUNG wire#w1
   RUNG wire#w1
      { S7_Templates := "SrcType := Real" } EQ_Contact(in1 := #HMI_SPEED, in2 := 0.0)
      wire#w2
      Move(in := 10.0, out1 => #HMI_SPEED)
   END_RUNG
   RUNG wire#w1
      { S7_Templates := "SrcType := Int" } EQ_Contact(in1 := #STEP_85, in2 := #SQCR)
   END_RUNG wire#w2
   RUNG wire#w1
      { S7_Templates := "SrcType := Int" } EQ_Contact(in1 := #STEP_55, in2 := #SQCR)
      Move(in := 2.0, out1 => #HMI_SPEED)
   END_RUNG
   RUNG wire#powerrail
      Contact( "LOG_0" )
      Coil( #CONTROL_AUTOMAT.B2 )
   END_RUNG
   // the same network as SCL:
   #CONTROL_AUTOMAT.B3 := (#STEP_10 = #SQCR) OR ((#STEP_10 <= #SQCR) AND (#STEP_30 >= #SQCR)) OR (#STEP_45 = #SQCR) OR (#STEP_55 = #SQCR) OR (#STEP_85 = #SQCR);
   IF #CONTROL_AUTOMAT.B3 AND ((#HMI_SPEED = 0.0) OR (#STEP_85 = #SQCR)) THEN #HMI_SPEED := 10.0; END_IF;
   IF #CONTROL_AUTOMAT.B3 AND (#STEP_55 = #SQCR) THEN #HMI_SPEED := 2.0; END_IF;
   #CONTROL_AUTOMAT.B2 := "LOG_0";
END_REGION

REGION Network 24: automa DVERE / automa ARETOVANI
   RUNG wire#powerrail
      { S7_Templates := "SrcType := Int" } EQ_Contact(in1 := #STEP_50, in2 := #SQCR)
      Coil( #CONTROL_AUTOMAT.B4 )
   END_RUNG
   RUNG wire#powerrail
      { S7_Templates := "SrcType := Int" } EQ_Contact(in1 := #STEP_80, in2 := #SQCR)
      wire#w1
      Coil( #CONTROL_AUTOMAT.B5 )
   END_RUNG
   RUNG wire#powerrail
      { S7_Templates := "SrcType := Int" } EQ_Contact(in1 := #STEP_1005_START_INICIAL, in2 := #SQCR)
   END_RUNG wire#w1
   // the same network as SCL:
   #CONTROL_AUTOMAT.B4 := #STEP_50 = #SQCR;
   #CONTROL_AUTOMAT.B5 := (#STEP_80 = #SQCR) OR (#STEP_1005_START_INICIAL = #SQCR);
END_REGION

REGION Network 25: CONTROL BLOCK podavač / CONTROL BLOCK DVERE
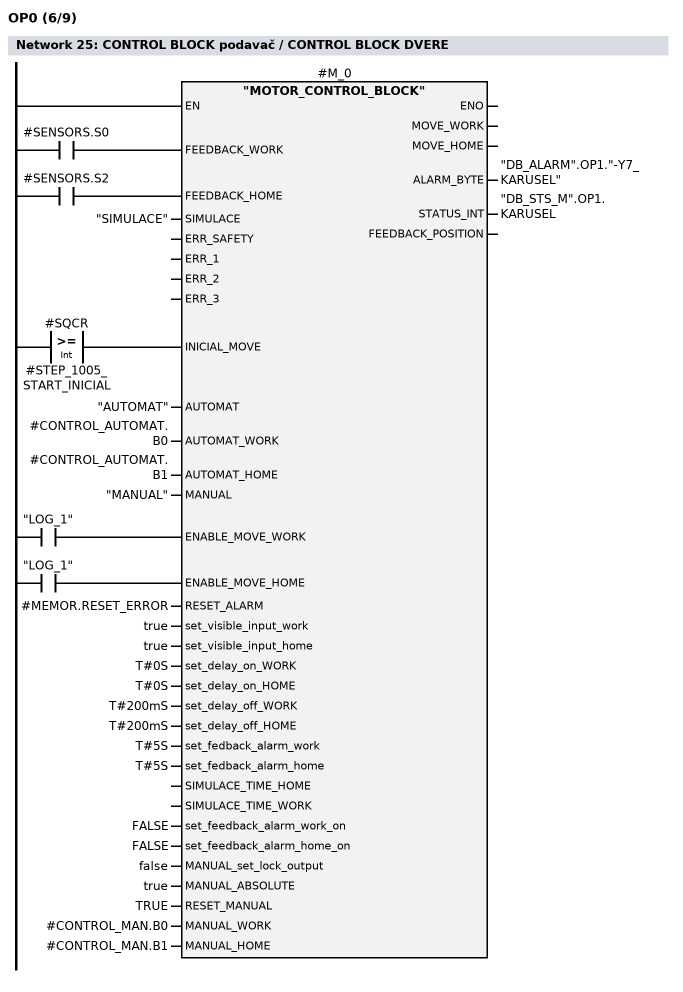
   RUNG wire#powerrail
      #M_0(FEEDBACK_WORK := wire#w1, FEEDBACK_HOME := wire#w2, INICIAL_MOVE := wire#w3, ENABLE_MOVE_WORK := wire#w4, ENABLE_MOVE_HOME := wire#w5, SIMULACE := "SIMULACE", ERR_SAFETY :=, ERR_1 :=, ERR_2 :=, ERR_3 :=, AUTOMAT := "AUTOMAT", AUTOMAT_WORK := #CONTROL_AUTOMAT.B0, AUTOMAT_HOME := #CONTROL_AUTOMAT.B1, MANUAL := "MANUAL", RESET_ALARM := #MEMOR.RESET_ERROR, set_visible_input_work := true, set_visible_input_home := true, set_delay_on_WORK := T#0S, set_delay_on_HOME := T#0S, set_delay_off_WORK := T#200mS, set_delay_off_HOME := T#200mS, set_fedback_alarm_work := T#5S, set_fedback_alarm_home := T#5S, SIMULACE_TIME_HOME :=, SIMULACE_TIME_WORK :=, set_feedback_alarm_work_on := FALSE, set_feedback_alarm_home_on := FALSE, MANUAL_set_lock_output := false, MANUAL_ABSOLUTE := true, RESET_MANUAL := TRUE, MANUAL_WORK := #CONTROL_MAN.B0, MANUAL_HOME := #CONTROL_MAN.B1, MOVE_WORK =>, MOVE_HOME =>, ALARM_BYTE => "DB_ALARM".OP1."-Y7_KARUSEL", STATUS_INT => "DB_STS_M".OP1.KARUSEL, FEEDBACK_POSITION =>)
   END_RUNG
   RUNG wire#powerrail
      Contact( #SENSORS.S0 )
   END_RUNG wire#w1
   RUNG wire#powerrail
      Contact( #SENSORS.S2 )
   END_RUNG wire#w2
   RUNG wire#powerrail
      { S7_Templates := "SrcType := Int" } GE_Contact(in1 := #SQCR, in2 := #STEP_1005_START_INICIAL)
   END_RUNG wire#w3
   RUNG wire#powerrail
      Contact( "LOG_1" )
   END_RUNG wire#w4
   RUNG wire#powerrail
      Contact( "LOG_1" )
   END_RUNG wire#w5
   // the same network as SCL:
   #M_0(FEEDBACK_WORK := #SENSORS.S0,   // "MOTOR_CONTROL_BLOCK"
        FEEDBACK_HOME := #SENSORS.S2,
        SIMULACE := "SIMULACE",
        INICIAL_MOVE := #SQCR >= #STEP_1005_START_INICIAL,
        AUTOMAT := "AUTOMAT",
        AUTOMAT_WORK := #CONTROL_AUTOMAT.B0,
        AUTOMAT_HOME := #CONTROL_AUTOMAT.B1,
        MANUAL := "MANUAL",
        ENABLE_MOVE_WORK := "LOG_1",
        ENABLE_MOVE_HOME := "LOG_1",
        RESET_ALARM := #MEMOR.RESET_ERROR,
        set_visible_input_work := true,
        set_visible_input_home := true,
        set_delay_on_WORK := T#0S,
        set_delay_on_HOME := T#0S,
        set_delay_off_WORK := T#200mS,
        set_delay_off_HOME := T#200mS,
        set_fedback_alarm_work := T#5S,
        set_fedback_alarm_home := T#5S,
        set_feedback_alarm_work_on := FALSE,
        set_feedback_alarm_home_on := FALSE,
        MANUAL_set_lock_output := false,
        MANUAL_ABSOLUTE := true,
        RESET_MANUAL := TRUE,
        MANUAL_WORK := #CONTROL_MAN.B0,
        MANUAL_HOME := #CONTROL_MAN.B1,
        ALARM_BYTE => "DB_ALARM".OP1."-Y7_KARUSEL",
        STATUS_INT => "DB_STS_M".OP1.KARUSEL);
END_REGION

REGION Network 26: CONTROL BLOCK dopravník / CONTROL BLOCK OSA Z
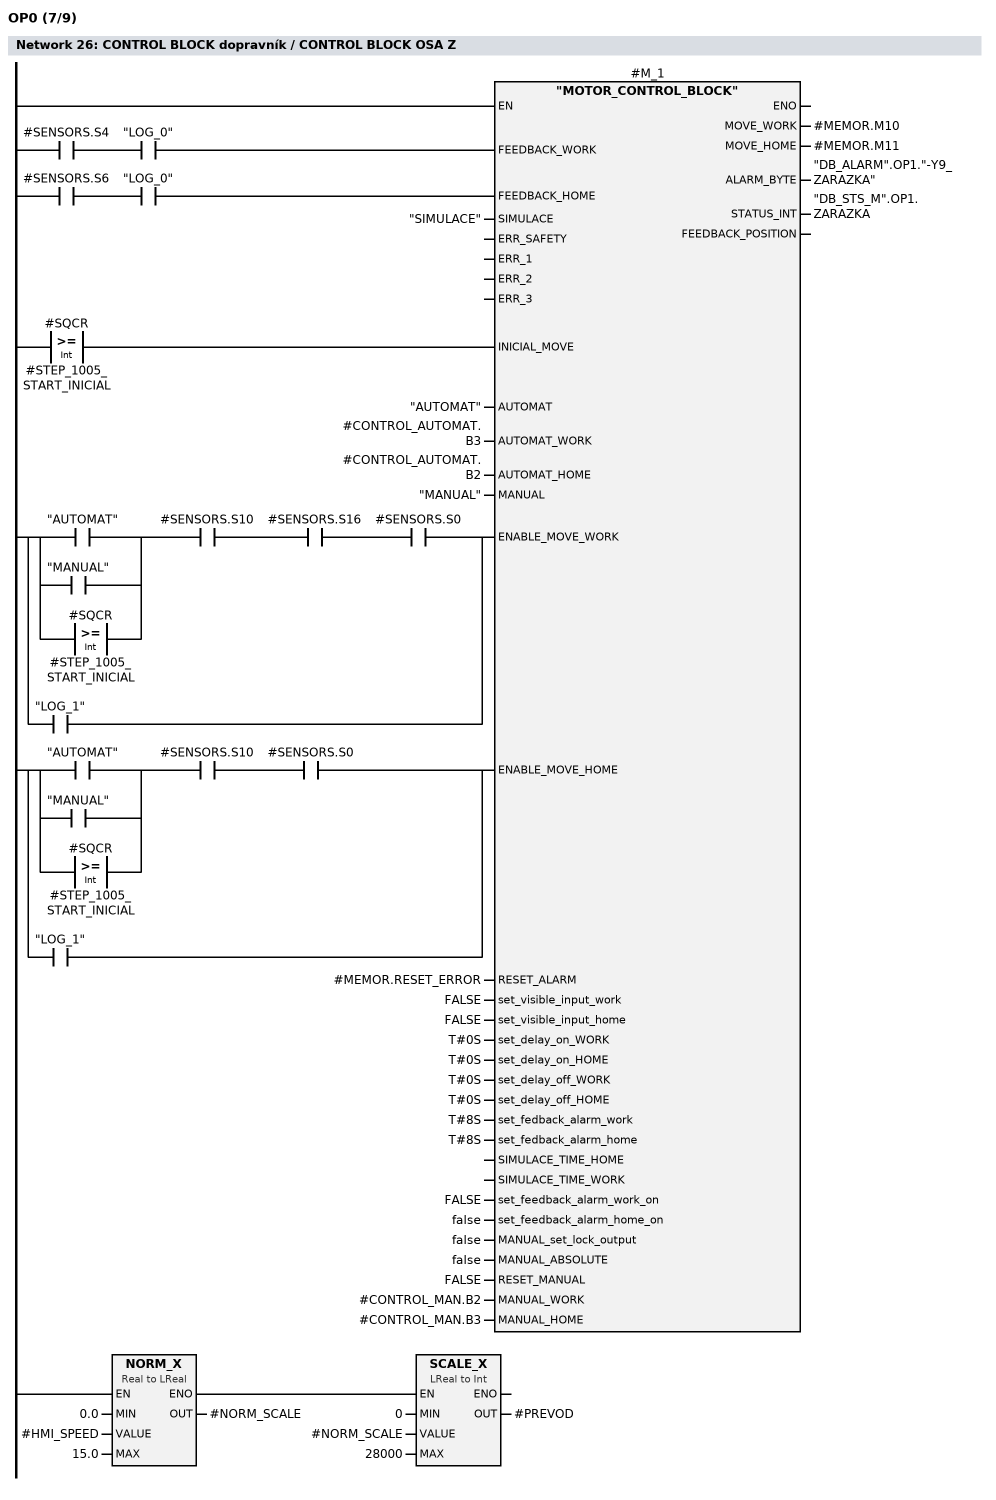
   RUNG wire#powerrail
      #M_1(FEEDBACK_WORK := wire#w1, FEEDBACK_HOME := wire#w2, INICIAL_MOVE := wire#w3, ENABLE_MOVE_WORK := wire#w5, ENABLE_MOVE_HOME := wire#w7, SIMULACE := "SIMULACE", ERR_SAFETY :=, ERR_1 :=, ERR_2 :=, ERR_3 :=, AUTOMAT := "AUTOMAT", AUTOMAT_WORK := #CONTROL_AUTOMAT.B3, AUTOMAT_HOME := #CONTROL_AUTOMAT.B2, MANUAL := "MANUAL", RESET_ALARM := #MEMOR.RESET_ERROR, set_visible_input_work := FALSE, set_visible_input_home := FALSE, set_delay_on_WORK := T#0S, set_delay_on_HOME := T#0S, set_delay_off_WORK := T#0S, set_delay_off_HOME := T#0S, set_fedback_alarm_work := T#8S, set_fedback_alarm_home := T#8S, SIMULACE_TIME_HOME :=, SIMULACE_TIME_WORK :=, set_feedback_alarm_work_on := FALSE, set_feedback_alarm_home_on := false, MANUAL_set_lock_output := false, MANUAL_ABSOLUTE := false, RESET_MANUAL := FALSE, MANUAL_WORK := #CONTROL_MAN.B2, MANUAL_HOME := #CONTROL_MAN.B3, MOVE_WORK => #MEMOR.M10, MOVE_HOME => #MEMOR.M11, ALARM_BYTE => "DB_ALARM".OP1."-Y9_ZARAZKA", STATUS_INT => "DB_STS_M".OP1.ZARAZKA, FEEDBACK_POSITION =>)
   END_RUNG
   RUNG wire#powerrail
      Contact( #SENSORS.S4 )
      Contact( "LOG_0" )
   END_RUNG wire#w1
   RUNG wire#powerrail
      Contact( #SENSORS.S6 )
      Contact( "LOG_0" )
   END_RUNG wire#w2
   RUNG wire#powerrail
      { S7_Templates := "SrcType := Int" } GE_Contact(in1 := #SQCR, in2 := #STEP_1005_START_INICIAL)
   END_RUNG wire#w3
   RUNG wire#powerrail
      Contact( "AUTOMAT" )
      wire#w4
      Contact( #SENSORS.S10 )
      Contact( #SENSORS.S16 )
      Contact( #SENSORS.S0 )
   END_RUNG wire#w5
   RUNG wire#powerrail
      Contact( "MANUAL" )
   END_RUNG wire#w4
   RUNG wire#powerrail
      { S7_Templates := "SrcType := Int" } GE_Contact(in1 := #SQCR, in2 := #STEP_1005_START_INICIAL)
   END_RUNG wire#w4
   RUNG wire#powerrail
      Contact( "LOG_1" )
   END_RUNG wire#w5
   RUNG wire#powerrail
      Contact( "AUTOMAT" )
      wire#w6
      Contact( #SENSORS.S10 )
      Contact( #SENSORS.S0 )
   END_RUNG wire#w7
   RUNG wire#powerrail
      Contact( "MANUAL" )
   END_RUNG wire#w6
   RUNG wire#powerrail
      { S7_Templates := "SrcType := Int" } GE_Contact(in1 := #SQCR, in2 := #STEP_1005_START_INICIAL)
   END_RUNG wire#w6
   RUNG wire#powerrail
      Contact( "LOG_1" )
   END_RUNG wire#w7
   RUNG wire#powerrail
      { S7_Templates := "[SrcType := Real, DestType := LReal]" } Normalize(min := 0.0, value := #HMI_SPEED, max := 15.0, out => #NORM_SCALE)
      { S7_Templates := "[SrcType := LReal, DestType := Int]" } Scale(min := 0, value := #NORM_SCALE, max := 28000, out => #PREVOD)
   END_RUNG
   // the same network as SCL:
   #M_1(FEEDBACK_WORK := #SENSORS.S4 AND "LOG_0",   // "MOTOR_CONTROL_BLOCK"
        FEEDBACK_HOME := #SENSORS.S6 AND "LOG_0",
        SIMULACE := "SIMULACE",
        INICIAL_MOVE := #SQCR >= #STEP_1005_START_INICIAL,
        AUTOMAT := "AUTOMAT",
        AUTOMAT_WORK := #CONTROL_AUTOMAT.B3,
        AUTOMAT_HOME := #CONTROL_AUTOMAT.B2,
        MANUAL := "MANUAL",
        ENABLE_MOVE_WORK := (("AUTOMAT" OR "MANUAL" OR (#SQCR >= #STEP_1005_START_INICIAL)) AND #SENSORS.S10 AND #SENSORS.S16 AND #SENSORS.S0) OR "LOG_1",
        ENABLE_MOVE_HOME := (("AUTOMAT" OR "MANUAL" OR (#SQCR >= #STEP_1005_START_INICIAL)) AND #SENSORS.S10 AND #SENSORS.S0) OR "LOG_1",
        RESET_ALARM := #MEMOR.RESET_ERROR,
        set_visible_input_work := FALSE,
        set_visible_input_home := FALSE,
        set_delay_on_WORK := T#0S,
        set_delay_on_HOME := T#0S,
        set_delay_off_WORK := T#0S,
        set_delay_off_HOME := T#0S,
        set_fedback_alarm_work := T#8S,
        set_fedback_alarm_home := T#8S,
        set_feedback_alarm_work_on := FALSE,
        set_feedback_alarm_home_on := false,
        MANUAL_set_lock_output := false,
        MANUAL_ABSOLUTE := false,
        RESET_MANUAL := FALSE,
        MANUAL_WORK := #CONTROL_MAN.B2,
        MANUAL_HOME := #CONTROL_MAN.B3,
        MOVE_WORK => #MEMOR.M10,
        MOVE_HOME => #MEMOR.M11,
        ALARM_BYTE => "DB_ALARM".OP1."-Y9_ZARAZKA",
        STATUS_INT => "DB_STS_M".OP1.ZARAZKA);
   #NORM_SCALE := NORM_X(MIN := 0.0, VALUE := #HMI_SPEED, MAX := 15.0);
   #PREVOD := SCALE_X(MIN := 0, VALUE := #NORM_SCALE, MAX := 28000);
END_REGION

REGION Network 27: CONTROL BLOCK dveře laser / CONTROL BLOCK ARETACE HLAVY
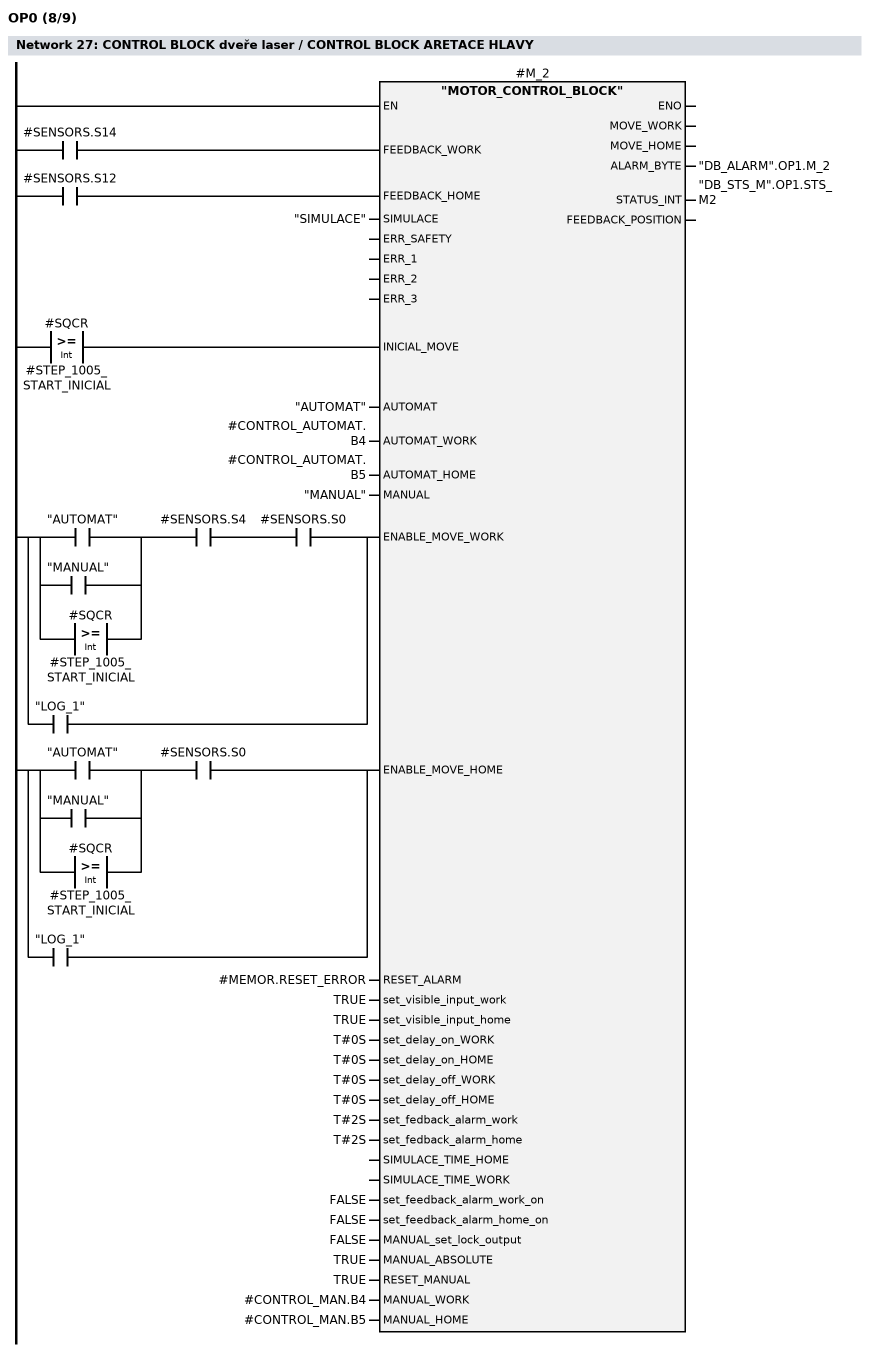
   RUNG wire#powerrail
      #M_2(FEEDBACK_WORK := wire#w1, FEEDBACK_HOME := wire#w2, INICIAL_MOVE := wire#w3, ENABLE_MOVE_WORK := wire#w5, ENABLE_MOVE_HOME := wire#w7, SIMULACE := "SIMULACE", ERR_SAFETY :=, ERR_1 :=, ERR_2 :=, ERR_3 :=, AUTOMAT := "AUTOMAT", AUTOMAT_WORK := #CONTROL_AUTOMAT.B4, AUTOMAT_HOME := #CONTROL_AUTOMAT.B5, MANUAL := "MANUAL", RESET_ALARM := #MEMOR.RESET_ERROR, set_visible_input_work := TRUE, set_visible_input_home := TRUE, set_delay_on_WORK := T#0S, set_delay_on_HOME := T#0S, set_delay_off_WORK := T#0S, set_delay_off_HOME := T#0S, set_fedback_alarm_work := T#2S, set_fedback_alarm_home := T#2S, SIMULACE_TIME_HOME :=, SIMULACE_TIME_WORK :=, set_feedback_alarm_work_on := FALSE, set_feedback_alarm_home_on := FALSE, MANUAL_set_lock_output := FALSE, MANUAL_ABSOLUTE := TRUE, RESET_MANUAL := TRUE, MANUAL_WORK := #CONTROL_MAN.B4, MANUAL_HOME := #CONTROL_MAN.B5, MOVE_WORK =>, MOVE_HOME =>, ALARM_BYTE => "DB_ALARM".OP1.M_2, STATUS_INT => "DB_STS_M".OP1.STS_M2, FEEDBACK_POSITION =>)
   END_RUNG
   RUNG wire#powerrail
      Contact( #SENSORS.S14 )
   END_RUNG wire#w1
   RUNG wire#powerrail
      Contact( #SENSORS.S12 )
   END_RUNG wire#w2
   RUNG wire#powerrail
      { S7_Templates := "SrcType := Int" } GE_Contact(in1 := #SQCR, in2 := #STEP_1005_START_INICIAL)
   END_RUNG wire#w3
   RUNG wire#powerrail
      Contact( "AUTOMAT" )
      wire#w4
      Contact( #SENSORS.S4 )
      Contact( #SENSORS.S0 )
   END_RUNG wire#w5
   RUNG wire#powerrail
      Contact( "MANUAL" )
   END_RUNG wire#w4
   RUNG wire#powerrail
      { S7_Templates := "SrcType := Int" } GE_Contact(in1 := #SQCR, in2 := #STEP_1005_START_INICIAL)
   END_RUNG wire#w4
   RUNG wire#powerrail
      Contact( "LOG_1" )
   END_RUNG wire#w5
   RUNG wire#powerrail
      Contact( "AUTOMAT" )
      wire#w6
      Contact( #SENSORS.S0 )
   END_RUNG wire#w7
   RUNG wire#powerrail
      Contact( "MANUAL" )
   END_RUNG wire#w6
   RUNG wire#powerrail
      { S7_Templates := "SrcType := Int" } GE_Contact(in1 := #SQCR, in2 := #STEP_1005_START_INICIAL)
   END_RUNG wire#w6
   RUNG wire#powerrail
      Contact( "LOG_1" )
   END_RUNG wire#w7
   // the same network as SCL:
   #M_2(FEEDBACK_WORK := #SENSORS.S14,   // "MOTOR_CONTROL_BLOCK"
        FEEDBACK_HOME := #SENSORS.S12,
        SIMULACE := "SIMULACE",
        INICIAL_MOVE := #SQCR >= #STEP_1005_START_INICIAL,
        AUTOMAT := "AUTOMAT",
        AUTOMAT_WORK := #CONTROL_AUTOMAT.B4,
        AUTOMAT_HOME := #CONTROL_AUTOMAT.B5,
        MANUAL := "MANUAL",
        ENABLE_MOVE_WORK := (("AUTOMAT" OR "MANUAL" OR (#SQCR >= #STEP_1005_START_INICIAL)) AND #SENSORS.S4 AND #SENSORS.S0) OR "LOG_1",
        ENABLE_MOVE_HOME := (("AUTOMAT" OR "MANUAL" OR (#SQCR >= #STEP_1005_START_INICIAL)) AND #SENSORS.S0) OR "LOG_1",
        RESET_ALARM := #MEMOR.RESET_ERROR,
        set_visible_input_work := TRUE,
        set_visible_input_home := TRUE,
        set_delay_on_WORK := T#0S,
        set_delay_on_HOME := T#0S,
        set_delay_off_WORK := T#0S,
        set_delay_off_HOME := T#0S,
        set_fedback_alarm_work := T#2S,
        set_fedback_alarm_home := T#2S,
        set_feedback_alarm_work_on := FALSE,
        set_feedback_alarm_home_on := FALSE,
        MANUAL_set_lock_output := FALSE,
        MANUAL_ABSOLUTE := TRUE,
        RESET_MANUAL := TRUE,
        MANUAL_WORK := #CONTROL_MAN.B4,
        MANUAL_HOME := #CONTROL_MAN.B5,
        ALARM_BYTE => "DB_ALARM".OP1.M_2,
        STATUS_INT => "DB_STS_M".OP1.STS_M2);
END_REGION

REGION Network 28: EXTERNAL_TRIGER
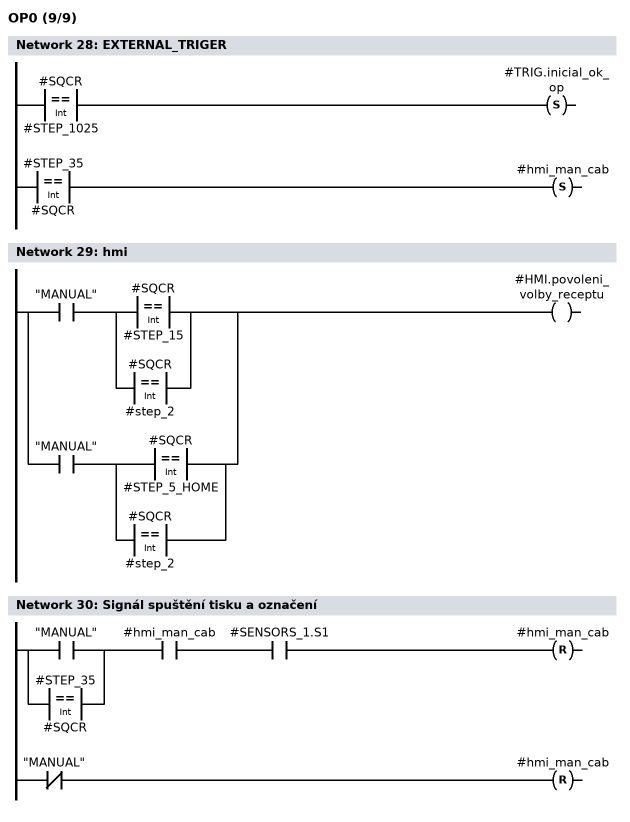
   RUNG wire#powerrail
      { S7_Templates := "SrcType := Int" } EQ_Contact(in1 := #SQCR, in2 := #STEP_1025)
      S_Coil( #TRIG.inicial_ok_op )
   END_RUNG
   RUNG wire#powerrail
      { S7_Templates := "SrcType := Int" } EQ_Contact(in1 := #STEP_35, in2 := #SQCR)
      S_Coil( #hmi_man_cab )
   END_RUNG
   // the same network as SCL:
   IF #SQCR = #STEP_1025 THEN #TRIG.inicial_ok_op := TRUE; END_IF;
   IF #STEP_35 = #SQCR THEN #hmi_man_cab := TRUE; END_IF;
END_REGION

REGION Network 29: hmi
   RUNG wire#powerrail
      Contact( "MANUAL" )
      wire#w1
      { S7_Templates := "SrcType := Int" } EQ_Contact(in1 := #SQCR, in2 := #STEP_15)
      wire#w2
      Coil( #HMI.povoleni_volby_receptu )
   END_RUNG
   RUNG wire#w1
      { S7_Templates := "SrcType := Int" } EQ_Contact(in1 := #SQCR, in2 := #step_2)
   END_RUNG wire#w2
   RUNG wire#powerrail
      Contact( "MANUAL" )
      wire#w3
      { S7_Templates := "SrcType := Int" } EQ_Contact(in1 := #SQCR, in2 := #STEP_5_HOME)
   END_RUNG wire#w2
   RUNG wire#w3
      { S7_Templates := "SrcType := Int" } EQ_Contact(in1 := #SQCR, in2 := #step_2)
   END_RUNG wire#w2
   // the same network as SCL:
   #HMI.povoleni_volby_receptu := ("MANUAL" AND ((#SQCR = #STEP_15) OR (#SQCR = #step_2))) OR ("MANUAL" AND ((#SQCR = #STEP_5_HOME) OR (#SQCR = #step_2)));
END_REGION

REGION Network 30: Signál spuštění tisku a označení
   RUNG wire#powerrail
      Contact( "MANUAL" )
      wire#w1
      Contact( #hmi_man_cab )
      Contact( #SENSORS_1.S1 )
      R_Coil( #hmi_man_cab )
   END_RUNG
   RUNG wire#powerrail
      { S7_Templates := "SrcType := Int" } EQ_Contact(in1 := #STEP_35, in2 := #SQCR)
   END_RUNG wire#w1
   RUNG wire#powerrail
      I_Contact( "MANUAL" )
      R_Coil( #hmi_man_cab )
   END_RUNG
   // the same network as SCL:
   IF ("MANUAL" OR (#STEP_35 = #SQCR)) AND #hmi_man_cab AND #SENSORS_1.S1 THEN #hmi_man_cab := FALSE; END_IF;
   IF NOT "MANUAL" THEN #hmi_man_cab := FALSE; END_IF;
END_REGION
END_FUNCTION_BLOCK

FUNCTION_BLOCK "OP1"   // FB50, LAD
{ S7_Optimized_Access := 'TRUE' }
VERSION : 0.1
   VAR
      CONTROL_MAN : Struct
         kar_work : Bool;
         kar_home : Bool;
         zarazka_work : Bool;
         zarazka_home : Bool;
         B4 : Bool;
         B5 : Bool;
         B6 : Bool;
         B7 : Bool;
         B8 : Bool;
         B9 : Bool;
         odfuk_1 : Bool;
         odfuk_2 : Bool;
         B12 : Bool;
         B13 : Bool;
         B14 : Bool;
         B15 : Bool;
         B16 : Bool;
         B17 : Bool;
         B18 : Bool;
         B19 : Bool;
         B20 : Bool;
         B21 : Bool;
         B22 : Bool;
         B23 : Bool;
         B24 : Bool;
         B25 : Bool;
         B26 : Bool;
         B27 : Bool;
         B28 : Bool;
         B29 : Bool;
         B30 : Bool;
         B31 : Bool;
      END_STRUCT;
      CONTROL_AUTOMAT : Struct
         KAR_WORK : Bool;
         KAR_HOME : Bool;
         ZARAZKA_WORK : Bool;
         ZARAZKA_HOME : Bool;
         B4 : Bool;
         B5 : Bool;
         B6 : Bool;
         B7 : Bool;
         B8 : Bool;
         B9 : Bool;
         odfuk_1 : Bool;
         odfuk_2 : Bool;
         B12 : Bool;
         B13 : Bool;
         B14 : Bool;
         B15 : Bool;
         B16 : Bool;
         B17 : Bool;
         B18 : Bool;
         B19 : Bool;
         B20 : Bool;
         B21 : Bool;
         B22 : Bool;
         B23 : Bool;
         B24 : Bool;
         B25 : Bool;
         B26 : Bool;
         B27 : Bool;
         B28 : Bool;
         B29 : Bool;
         B30 : Bool;
         B31 : Bool;
      END_STRUCT;
      SENSORS : Struct
         prechod_1 : Bool;
         prechod_1_neg : Bool;
         kontrola : Bool;
         kontrola_neg : Bool;
         prechod_2 : Bool;
         Prechod_2_neg : Bool;
         Pozice_vyrazovace : Bool;
         Pozice_vyrazovace_neg : Bool;
         Pozice_pistu : Bool;   // KARUSEL JE NATOČEN PŘÍPRAVKEM A K BRÁNĚ
         Pozice_pistu_neg : Bool;
         s10 : Bool;
         s11 : Bool;
         s12 : Bool;
         s13 : Bool;
         s14 : Bool;
         s15 : Bool;
         s16 : Bool;
         s17 : Bool;
         s18 : Bool;
         s19 : Bool;
         s20 : Bool;
         s21 : Bool;
         s22 : Bool;
         s23 : Bool;
         s24 : Bool;
         s25 : Bool;
         s26 : Bool;
         s27 : Bool;
         s28 : Bool;
         s29 : Bool;
         s30 : Bool;
         s31 : Bool;
      END_STRUCT;
      SENSORS_1 : Struct
         S0 : Bool;
         S1 : Bool;
         S2 : Bool;
         S3 : Bool;
         S4 : Bool;
         S5 : Bool;
         S6 : Bool;
         S7 : Bool;
         S8 : Bool;
         S9 : Bool;
         SESTAVA_NENI_OTOCENA : Bool;
         SESTAVA_JE_OTOCENA : Bool;
         S12 : Bool;
         S13 : Bool;
         S14 : Bool;
         S15 : Bool;
         S16 : Bool;
         S17 : Bool;
         S18 : Bool;
         S19 : Bool;
         S20 : Bool;
         S21 : Bool;
         S22 : Bool;
         S23 : Bool;
         S24 : Bool;
         S25 : Bool;
         S26 : Bool;
         S27 : Bool;
         S28 : Bool;
         S29 : Bool;
         S30 : Bool;
         l_3_neg : Bool;
      END_STRUCT;
      S_0 : "SENSOR";
      S_1 : "SENSOR";
      S_2 : "SENSOR";
      S_3 : "SENSOR";
      S_4 : "SENSOR";
      S_5 : "SENSOR";
      S_6 : "SENSOR";
      M_karusel : "MOTOR_CONTROL_BLOCK";
      M_zarazka : "MOTOR_CONTROL_BLOCK";
      M_CLONA : "MOTOR_CONTROL_BLOCK";
      SQCR : Int;
      hmi_sqcr : Int;
      TRIG : Struct
         inicial_ok_op : Bool;
         DSSAD : Bool;
         INICIALIZACE_PROBEHLA : Bool;
         trig_dil : Bool;
         p_trig_control_tcon : Bool;
         T6 : Bool;
         SPUST_OP_4 : Bool;
         vlez_do_zavory_pri_rotaci : Bool;
         START_INICIAL_OP2 : Bool;
         START_INICIAL_OP3 : Bool;
         spust_odsavani : Bool;
         VYPRAZNI_OK_OP_2_A : Bool;
         VYPRAZNI_NOK_OP_2_A : Bool;
         VYPRAZDNI_OK_OP_3_B : Bool;
         VYPRAZDNI_NOK_OP_3_B : Bool;
         RESET_NCODER : Bool;
         op_1_ready : Bool;
      END_STRUCT;
      MEMOR : Struct
         n_trig_vypnuti : Bool;
         M1 : Bool;
         M2 : Bool;
         M3 : Bool;
         M4 : Bool;
         p_trig_odavacka : Bool;
         M6 : Bool;
         M7 : Bool;
         M8 : Bool;
         M9 : Bool;
         M10 : Bool;
         M11 : Bool;
         RESET_ERROR : Bool;
         vyrazeni_pamet : Bool;
         M14 : Bool;
         M15 : Bool;
         SETOVANI_START : Bool;
         M17 : Bool;
         p_trig_pamet_1 : Bool;
         p_trig_pamet_2 : Bool;
         p_trig_pamet_3 : Bool;
         p_trig_pamet_4 : Bool;
         p_trig_pamet_5 : Bool;
         p_trig_pamet_6 : Bool;
         p_trig_pamet_7 : Bool;
         p_trig_pamet_8 : Bool;
         p_trig_pamet_9 : Bool;
         p_trig_pamet_10 : Bool;
         p_trig_vyrad : Bool;
         p_Trig_cisteni_pozice : Bool;
         p_trig_citac : Bool;
         N_TRIG_SAFETY : Bool;
         P_TRIG_RESET_POZICE : Bool;
         M33 : Bool;
         start_caklu : Bool;
         M35 : Bool;
         M36 : Bool;
         M37 : Bool;
         M38 : Bool;
         M39 : Bool;
         ALARM_GLOBAL : Bool;
         M41 : Bool;
         M42 : Bool;
         M43 : Bool;
         M44 : Bool;
         M45 : Bool;
         M46 : Bool;
         M47 : Bool;
         M48 : Bool;
         M49 : Bool;
         wrong_p_trig : Bool;
         alarm_p_trig : Bool;
         M52 : Bool;
         M53 : Bool;
         M54 : Bool;
         M55 : Bool;
         M56 : Bool;
         M57 : Bool;
         M58 : Bool;
         M59 : Bool;
         M60 : Bool;
         M61 : Bool;
         M62 : Bool;
         M63 : Bool;
      END_STRUCT;
      "TIMER" : Struct
         TIMER_0 : IEC_TIMER;
         TIMER_VACUUM_CLEANER : IEC_TIMER;
         TIMER_DELAY_RESET_EXECUTE : IEC_TIMER;
         TIMER_3 : IEC_TIMER;
         TIMER_4 : IEC_TIMER;
         air : IEC_TIMER;
         TIMER_6 : IEC_TIMER;
         TIMER_7 : IEC_TIMER;
      END_STRUCT;
      HMI : Struct
         povoleni_volby_receptu : Bool;
         "svetlo_on/off" : Bool;
         ALARM_VIDITELNOST : Bool;
         hmi_3 : Bool;
         hmi_4 : Bool;
         reset_fronty : Bool;
         hmi_6 : Bool;
         hmi_7 : Bool;
         hmi_8 : Bool;
         hmi_9 : Bool;
         hmi_10 : Bool;
         hmi_11 : Bool;
         hmi_12 : Bool;
         hmi_13 : Bool;
         hmi_14 : Bool;
         hmi_15 : Bool;
      END_STRUCT;
      STRING_0 : String[1];
      array_chyb_ctec : Array[1..16] of Bool;
      zpracovani_dat : Array[1..1] of Struct
         prenaseny_text : String[100];
         balik_den : Int;
         vyrazeni : Bool;
      END_STRUCT;
      aktual_kusy : Int;
      i : Int;
      q : Int;
      pocet_znaku_string_kamera : Int;
      ocekavany_text : String[100];
      format_etiketa_ok : Bool;
      Kamera : Struct
         s2_pamet : Bool;
         s2_nabeh : Bool;
         sber_aktivni : Bool;
         prijato_etiketa : Bool;
         prijato_folie_l : Bool;
         prijato_folie_p : Bool;
         ok_etiketa : Bool;
         ok_folie_l : Bool;
         ok_folie_p : Bool;
         vyradit : Bool;
         fronta_plna : Bool;   // alarm
         bypass_ocr : Bool := True;   // dočasně, dokud není doladěné OCR
         last_id_etiketa : Word;
         last_id_folie_l : Word;
         last_id_folie_p : Word;
         balik_den : Int;
         idx : Int;
         pocet : Int;
         text_etiketa : String[100];
         timeout_sberu : Time :=  T#1S;
         kontrola_tridirny : Bool := true;   // HMI: kontrola kódu třídírny zapnuta
         tridirna_ok : Bool;   // výsledek kontroly posledního plata (pro online diagnostiku)
      END_STRUCT;
      Vyrazeni : Struct
         s4_pamet : Bool;
         s4_nabeh : Bool;
         aktivni : Bool;
         vyradit : Bool;
         chyba_bez_dat : Bool;   // alarm: plato u vyřazovače bez záznamu
         chyba_pist : Bool;   // alarm: píst nevyjel / nebyl v home
         max_puls : Time := T#200MS;
         vyrazovac_pripojen : Bool := true;   // TRUE až bude signál od dodavatele
         alarm_nok_balik : Bool;   // NOK plato prošlo bez vyřazení
         posledni_nok_balik : Int;   // číslo plata pro obsluhu / HMI
         posledni_nok_text : String[100];   // co přečetla kamera
         pocet_nok : DInt;   // počítadlo NOK plat
         pocet_bez_dat : DInt;
         majak_tp : TP_TIME;   // prodlouzeni blikani majaku pri vzrazenii
         majak : Bool;
      END_STRUCT;
      Kam_Etiketa_Job : Struct
         krok : Int;   // 0 klid, 10 odeslat, 20 čekat, 30 ukončit handshake
         pozadovany : Int;   // job z receptury (PRG_CAM_etiketa)
         odesli_pamet : Bool;   // hrana ODESLI_dATA
         aktivni : Bool;   // probíhá načítání jobu → blokovat triggery
         chyba : Bool;   // alarm: job se nepodařilo načíst
         chyba_kod : Word;   // CommandResultCode při chybě
         nesouhlasi : Bool;   // alarm: job v kameře ≠ job z receptury
         timeout : Time := T#10S;   // max. doba načítání jobu
      END_STRUCT;
      Test_tp_ka12 : TP_TIME;
   END_VAR
   VAR_TEMP
      DATA : Array[0..255] of Char;
      ARRAY_NULL : Array[1..8] of Bool;
      array_null_fronta : Array[1..1] of Struct
         prenaseny_text : String[100];
         balik_den : Int;
         vyrazeni : Bool;
      END_STRUCT;
      "char" : Array[0..0] of Char;
      "string" : String;
      cas : DTL;
      ret : Int;
   END_VAR
   VAR CONSTANT
      STEP_0 : Int := 0;
      step_2 : Int := 2;
      STEP_4 : Int := 4;
      STEP_5_HOME : Int := 5;
      STEP_7 : Int := 7;
      STEP_10 : Int := 10;
      STEP_15 : Int := 15;
      STEP_20 : Int := 20;
      STEP_23 : Int := 23;
      STEP_25 : Int := 25;
      STEP_27 : Int := 27;
      STEP_30 : Int := 30;
      STEP_35 : Int := 35;
      STEP_37 : Int := 37;
      STEP_40 : Int := 40;
      STEP_45 : Int := 45;
      STEP_50 : Int := 50;
      STEP_55 : Int := 55;
      STEP_60 : Int := 60;
      STEP_65 : Int := 65;
      STEP_70 : Int := 70;
      STEP_75 : Int := 75;
      STEP_80 : Int := 80;
      STEP_83 : Int := 83;
      STEP_85 : Int := 85;
      STEP_90 : Int := 90;
      STEP_95 : Int := 95;
      STEP_100 : Int := 100;
      STEP_105 : Int := 105;
      STEP_110 : Int := 110;
      STEP_113 : Int := 113;
      STEP_115 : Int := 115;
      STEP_120 : Int := 120;
      STEP_125 : Int := 125;
      STEP_130 : Int := 130;
      STEP_135 : Int := 135;
      STEP_140 : Int := 140;
      STEP_145 : Int := 145;
      STEP_150 : Int := 150;
      STEP_155 : Int := 155;
      STEP_1000 : Int := 1000;
      STEP_1001 : Int := 1001;
      STEP_1002 : Int := 1002;
      STEP_1003 : Int := 1003;
      STEP_1004 : Int := 1004;
      STEP_1005 : Int := 1005;
      STEP_1010 : Int := 1010;
      STEP_1015 : Int := 1015;
      STEP_1020 : Int := 1020;
      STEP_1025 : Int := 1025;
      STEP_3000 : Int := 3000;
      STEP_3005 : Int := 3005;
      STEP_3010 : Int := 3010;
      STEP_3015 : Int := 3015;
      STEP_3020 : Int := 3020;
      STEP_2000 : Int := 2000;
      string_null : String;
      char_null : Char;
      text_kartacek : String := 'Kartacek';
      string_kar_A : String := 'A';
      string_kar_B : String := 'B';
      KOD_TRIDIRNY : String := 'CZ32880102';
   END_VAR
   VAR_TEMP   // added for the SCL form of the ladder/FBD networks
      _w1 : Bool;
      _w2 : Bool;
      _w3 : Bool;
   END_VAR
BEGIN

REGION Network 1: manuali ovladani reset
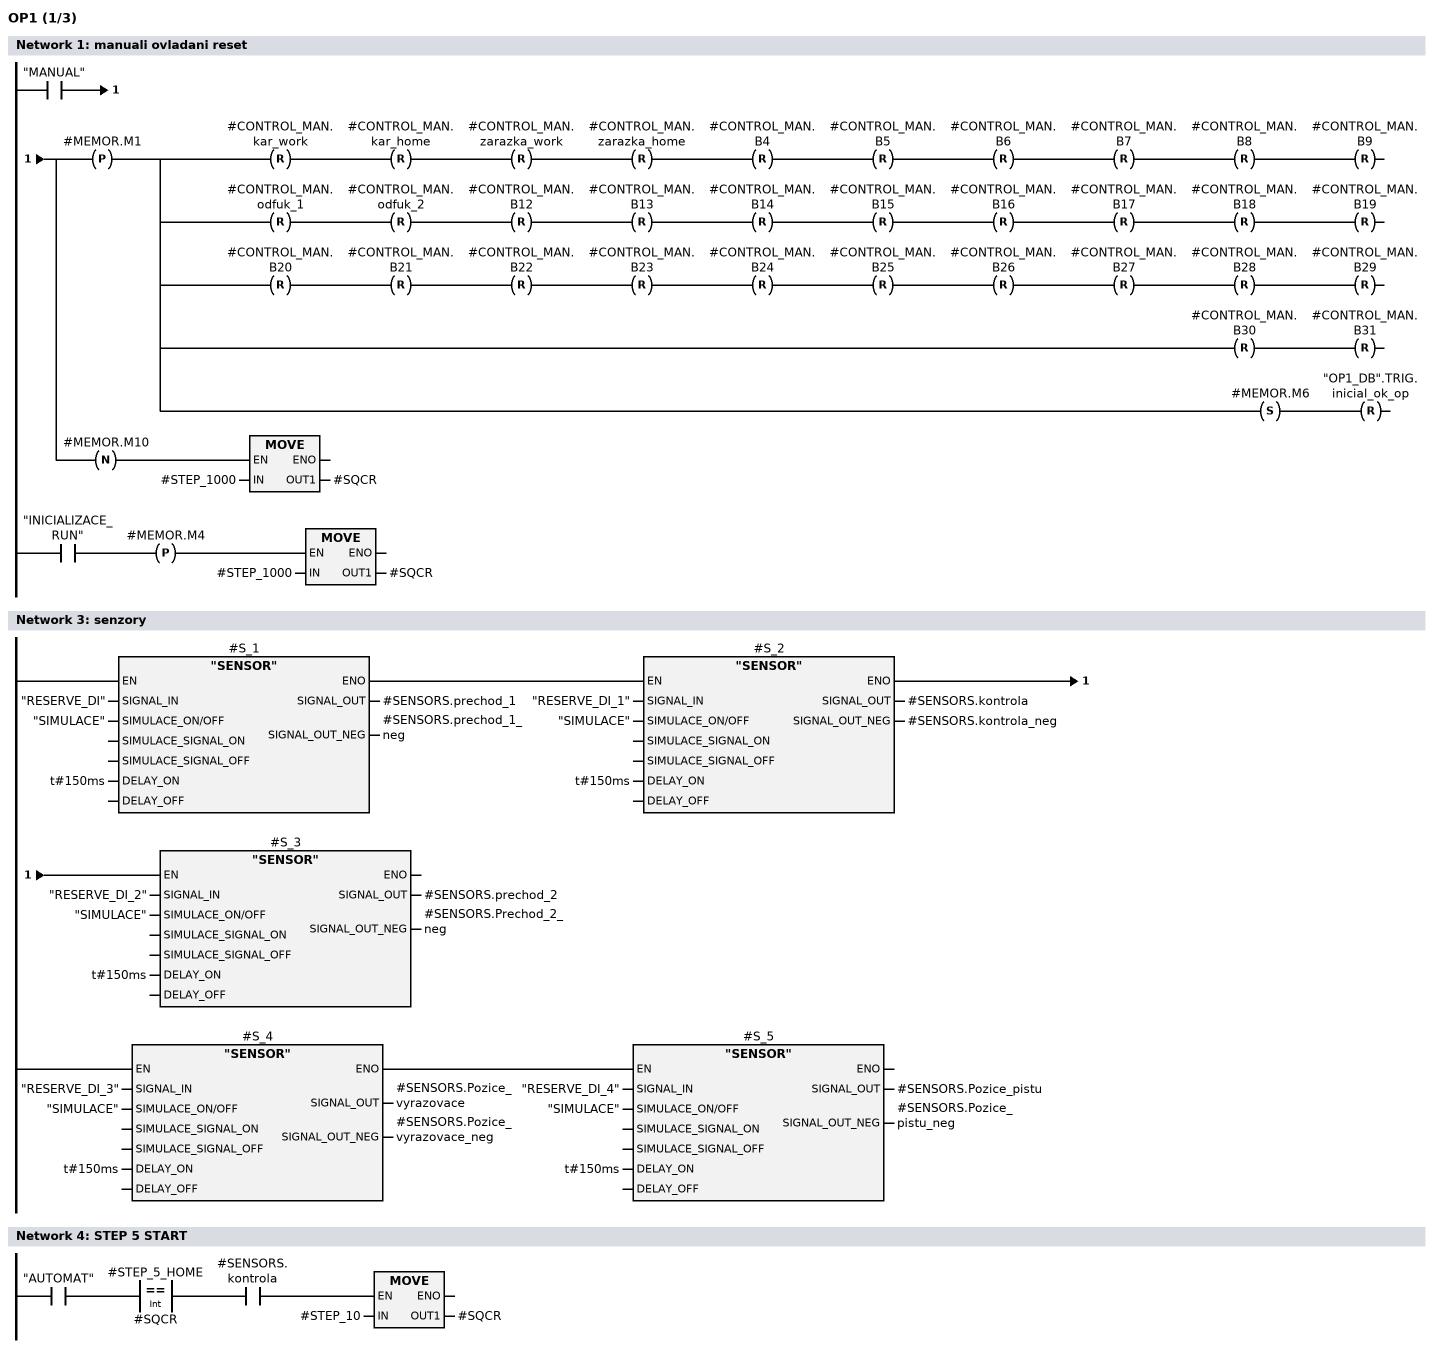
   RUNG wire#powerrail
      Contact( "MANUAL" )
      wire#w1
      P_Trig( #MEMOR.M1 )
      wire#w2
      R_Coil( #CONTROL_MAN.kar_work )
      R_Coil( #CONTROL_MAN.kar_home )
      R_Coil( #CONTROL_MAN.zarazka_work )
      R_Coil( #CONTROL_MAN.zarazka_home )
      R_Coil( #CONTROL_MAN.B4 )
      R_Coil( #CONTROL_MAN.B5 )
      R_Coil( #CONTROL_MAN.B6 )
      R_Coil( #CONTROL_MAN.B7 )
      R_Coil( #CONTROL_MAN.B8 )
      R_Coil( #CONTROL_MAN.B9 )
   END_RUNG
   RUNG wire#w2
      R_Coil( #CONTROL_MAN.odfuk_1 )
      R_Coil( #CONTROL_MAN.odfuk_2 )
      R_Coil( #CONTROL_MAN.B12 )
      R_Coil( #CONTROL_MAN.B13 )
      R_Coil( #CONTROL_MAN.B14 )
      R_Coil( #CONTROL_MAN.B15 )
      R_Coil( #CONTROL_MAN.B16 )
      R_Coil( #CONTROL_MAN.B17 )
      R_Coil( #CONTROL_MAN.B18 )
      R_Coil( #CONTROL_MAN.B19 )
   END_RUNG
   RUNG wire#w2
      R_Coil( #CONTROL_MAN.B20 )
      R_Coil( #CONTROL_MAN.B21 )
      R_Coil( #CONTROL_MAN.B22 )
      R_Coil( #CONTROL_MAN.B23 )
      R_Coil( #CONTROL_MAN.B24 )
      R_Coil( #CONTROL_MAN.B25 )
      R_Coil( #CONTROL_MAN.B26 )
      R_Coil( #CONTROL_MAN.B27 )
      R_Coil( #CONTROL_MAN.B28 )
      R_Coil( #CONTROL_MAN.B29 )
   END_RUNG
   RUNG wire#w2
      R_Coil( #CONTROL_MAN.B30 )
      R_Coil( #CONTROL_MAN.B31 )
   END_RUNG
   RUNG wire#w2
      S_Coil( #MEMOR.M6 )
      R_Coil( "OP1_DB".TRIG.inicial_ok_op )
   END_RUNG
   RUNG wire#w1
      N_Trig( #MEMOR.M10 )
      Move(in := #STEP_1000, out1 => #SQCR)
   END_RUNG
   RUNG wire#powerrail
      Contact( "INICIALIZACE_RUN" )
      P_Trig( #MEMOR.M4 )
      Move(in := #STEP_1000, out1 => #SQCR)
   END_RUNG
   // the same network as SCL:
   #_w1 := "MANUAL" AND NOT #MEMOR.M1;   // rising edge
   #MEMOR.M1 := "MANUAL";
   IF #_w1 THEN
       #CONTROL_MAN.kar_work := FALSE;
       #CONTROL_MAN.kar_home := FALSE;
       #CONTROL_MAN.zarazka_work := FALSE;
       #CONTROL_MAN.zarazka_home := FALSE;
       #CONTROL_MAN.B4 := FALSE;
       #CONTROL_MAN.B5 := FALSE;
       #CONTROL_MAN.B6 := FALSE;
       #CONTROL_MAN.B7 := FALSE;
       #CONTROL_MAN.B8 := FALSE;
       #CONTROL_MAN.B9 := FALSE;
       #CONTROL_MAN.odfuk_1 := FALSE;
       #CONTROL_MAN.odfuk_2 := FALSE;
       #CONTROL_MAN.B12 := FALSE;
       #CONTROL_MAN.B13 := FALSE;
       #CONTROL_MAN.B14 := FALSE;
       #CONTROL_MAN.B15 := FALSE;
       #CONTROL_MAN.B16 := FALSE;
       #CONTROL_MAN.B17 := FALSE;
       #CONTROL_MAN.B18 := FALSE;
       #CONTROL_MAN.B19 := FALSE;
       #CONTROL_MAN.B20 := FALSE;
       #CONTROL_MAN.B21 := FALSE;
       #CONTROL_MAN.B22 := FALSE;
       #CONTROL_MAN.B23 := FALSE;
       #CONTROL_MAN.B24 := FALSE;
       #CONTROL_MAN.B25 := FALSE;
       #CONTROL_MAN.B26 := FALSE;
       #CONTROL_MAN.B27 := FALSE;
       #CONTROL_MAN.B28 := FALSE;
       #CONTROL_MAN.B29 := FALSE;
       #CONTROL_MAN.B30 := FALSE;
       #CONTROL_MAN.B31 := FALSE;
       #MEMOR.M6 := TRUE;
       "OP1_DB".TRIG.inicial_ok_op := FALSE;
   END_IF;
   #_w2 := NOT "MANUAL" AND #MEMOR.M10;   // falling edge
   #MEMOR.M10 := "MANUAL";
   IF #_w2 THEN #SQCR := #STEP_1000; END_IF;
   #_w3 := "INICIALIZACE_RUN" AND NOT #MEMOR.M4;   // rising edge
   #MEMOR.M4 := "INICIALIZACE_RUN";
   IF #_w3 THEN #SQCR := #STEP_1000; END_IF;
END_REGION

REGION Network 2: alarmy
END_REGION

REGION Network 3: senzory
   RUNG wire#powerrail
      #S_1(SIGNAL_IN := "RESERVE_DI", "SIMULACE_ON/OFF" := "SIMULACE", SIMULACE_SIGNAL_ON :=, SIMULACE_SIGNAL_OFF :=, DELAY_ON := t#150ms, DELAY_OFF :=, SIGNAL_OUT => #SENSORS.prechod_1, SIGNAL_OUT_NEG => #SENSORS.prechod_1_neg)
      #S_2(SIGNAL_IN := "RESERVE_DI_1", "SIMULACE_ON/OFF" := "SIMULACE", SIMULACE_SIGNAL_ON :=, SIMULACE_SIGNAL_OFF :=, DELAY_ON := t#150ms, DELAY_OFF :=, SIGNAL_OUT => #SENSORS.kontrola, SIGNAL_OUT_NEG => #SENSORS.kontrola_neg)
      #S_3(SIGNAL_IN := "RESERVE_DI_2", "SIMULACE_ON/OFF" := "SIMULACE", SIMULACE_SIGNAL_ON :=, SIMULACE_SIGNAL_OFF :=, DELAY_ON := t#150ms, DELAY_OFF :=, SIGNAL_OUT => #SENSORS.prechod_2, SIGNAL_OUT_NEG => #SENSORS.Prechod_2_neg)
   END_RUNG
   RUNG wire#powerrail
      #S_4(SIGNAL_IN := "RESERVE_DI_3", "SIMULACE_ON/OFF" := "SIMULACE", SIMULACE_SIGNAL_ON :=, SIMULACE_SIGNAL_OFF :=, DELAY_ON := t#150ms, DELAY_OFF :=, SIGNAL_OUT => #SENSORS.Pozice_vyrazovace, SIGNAL_OUT_NEG => #SENSORS.Pozice_vyrazovace_neg)
      #S_5(SIGNAL_IN := "RESERVE_DI_4", "SIMULACE_ON/OFF" := "SIMULACE", SIMULACE_SIGNAL_ON :=, SIMULACE_SIGNAL_OFF :=, DELAY_ON := t#150ms, DELAY_OFF :=, SIGNAL_OUT => #SENSORS.Pozice_pistu, SIGNAL_OUT_NEG => #SENSORS.Pozice_pistu_neg)
   END_RUNG
   // the same network as SCL:
   #S_1(SIGNAL_IN := "RESERVE_DI",   // "SENSOR"
        "SIMULACE_ON/OFF" := "SIMULACE",
        DELAY_ON := t#150ms,
        SIGNAL_OUT => #SENSORS.prechod_1,
        SIGNAL_OUT_NEG => #SENSORS.prechod_1_neg,
        ENO => #_w1);
   #S_2(EN := #_w1,   // "SENSOR"
        SIGNAL_IN := "RESERVE_DI_1",
        "SIMULACE_ON/OFF" := "SIMULACE",
        DELAY_ON := t#150ms,
        SIGNAL_OUT => #SENSORS.kontrola,
        SIGNAL_OUT_NEG => #SENSORS.kontrola_neg,
        ENO => #_w2);
   IF #_w2 THEN
       #S_3(SIGNAL_IN := "RESERVE_DI_2",   // "SENSOR"
            "SIMULACE_ON/OFF" := "SIMULACE",
            DELAY_ON := t#150ms,
            SIGNAL_OUT => #SENSORS.prechod_2,
            SIGNAL_OUT_NEG => #SENSORS.Prechod_2_neg);
   END_IF;
   #S_4(SIGNAL_IN := "RESERVE_DI_3",   // "SENSOR"
        "SIMULACE_ON/OFF" := "SIMULACE",
        DELAY_ON := t#150ms,
        SIGNAL_OUT => #SENSORS.Pozice_vyrazovace,
        SIGNAL_OUT_NEG => #SENSORS.Pozice_vyrazovace_neg,
        ENO => #_w3);
   IF #_w3 THEN
       #S_5(SIGNAL_IN := "RESERVE_DI_4",   // "SENSOR"
            "SIMULACE_ON/OFF" := "SIMULACE",
            DELAY_ON := t#150ms,
            SIGNAL_OUT => #SENSORS.Pozice_pistu,
            SIGNAL_OUT_NEG => #SENSORS.Pozice_pistu_neg);
   END_IF;
END_REGION

REGION Network 4: STEP 5 START
   RUNG wire#powerrail
      Contact( "AUTOMAT" )
      { S7_Templates := "SrcType := Int" } EQ_Contact(in1 := #STEP_5_HOME, in2 := #SQCR)
      Contact( #SENSORS.kontrola )
      Move(in := #STEP_10, out1 => #SQCR)
   END_RUNG
   // the same network as SCL:
   IF "AUTOMAT" AND (#STEP_5_HOME = #SQCR) AND #SENSORS.kontrola THEN #SQCR := #STEP_10; END_IF;
END_REGION

REGION Network 5: STEP 10
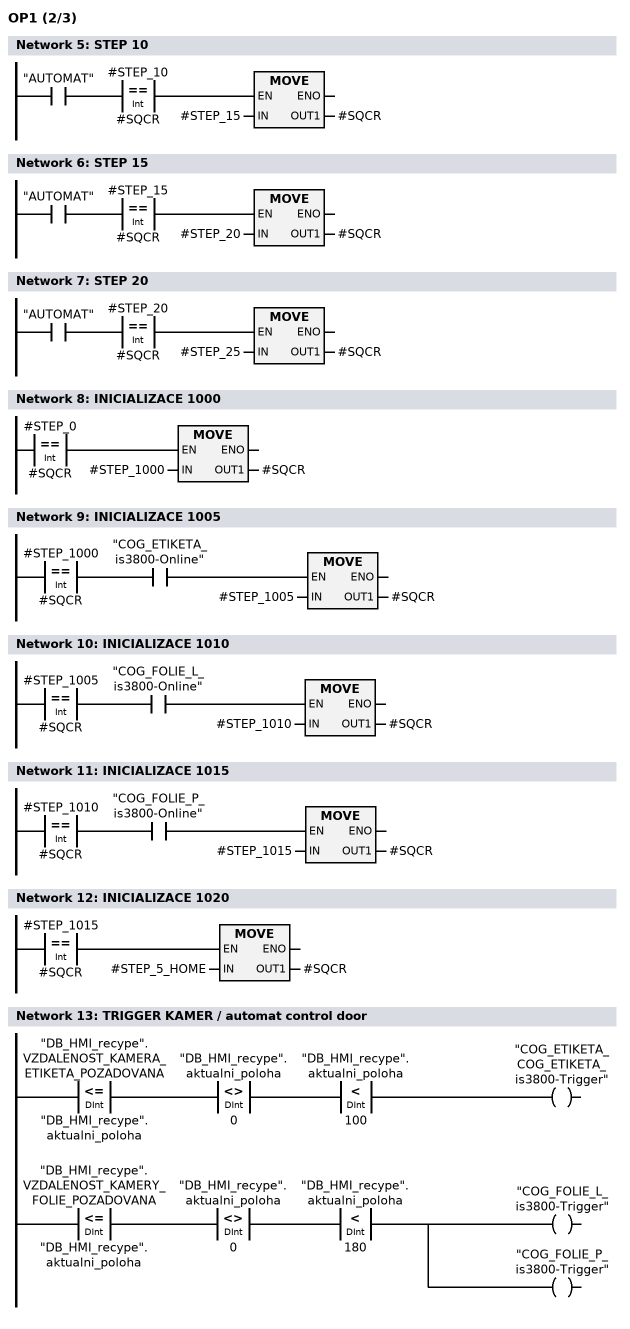
   RUNG wire#powerrail
      Contact( "AUTOMAT" )
      { S7_Templates := "SrcType := Int" } EQ_Contact(in1 := #STEP_10, in2 := #SQCR)
      Move(in := #STEP_15, out1 => #SQCR)
   END_RUNG
   // the same network as SCL:
   IF "AUTOMAT" AND (#STEP_10 = #SQCR) THEN #SQCR := #STEP_15; END_IF;
END_REGION

REGION Network 6: STEP 15
   RUNG wire#powerrail
      Contact( "AUTOMAT" )
      { S7_Templates := "SrcType := Int" } EQ_Contact(in1 := #STEP_15, in2 := #SQCR)
      Move(in := #STEP_20, out1 => #SQCR)
   END_RUNG
   // the same network as SCL:
   IF "AUTOMAT" AND (#STEP_15 = #SQCR) THEN #SQCR := #STEP_20; END_IF;
END_REGION

REGION Network 7: STEP 20
   RUNG wire#powerrail
      Contact( "AUTOMAT" )
      { S7_Templates := "SrcType := Int" } EQ_Contact(in1 := #STEP_20, in2 := #SQCR)
      Move(in := #STEP_25, out1 => #SQCR)
   END_RUNG
   // the same network as SCL:
   IF "AUTOMAT" AND (#STEP_20 = #SQCR) THEN #SQCR := #STEP_25; END_IF;
END_REGION

REGION Network 8: INICIALIZACE 1000
   RUNG wire#powerrail
      { S7_Templates := "SrcType := Int" } EQ_Contact(in1 := #STEP_0, in2 := #SQCR)
      Move(in := #STEP_1000, out1 => #SQCR)
   END_RUNG
   // the same network as SCL:
   IF #STEP_0 = #SQCR THEN #SQCR := #STEP_1000; END_IF;
END_REGION

REGION Network 9: INICIALIZACE 1005
   RUNG wire#powerrail
      { S7_Templates := "SrcType := Int" } EQ_Contact(in1 := #STEP_1000, in2 := #SQCR)
      Contact( "COG_ETIKETA_is3800-Online" )
      Move(in := #STEP_1005, out1 => #SQCR)
   END_RUNG
   // the same network as SCL:
   IF (#STEP_1000 = #SQCR) AND "COG_ETIKETA_is3800-Online" THEN #SQCR := #STEP_1005; END_IF;
END_REGION

REGION Network 10: INICIALIZACE 1010
   RUNG wire#powerrail
      { S7_Templates := "SrcType := Int" } EQ_Contact(in1 := #STEP_1005, in2 := #SQCR)
      Contact( "COG_FOLIE_L_is3800-Online" )
      Move(in := #STEP_1010, out1 => #SQCR)
   END_RUNG
   // the same network as SCL:
   IF (#STEP_1005 = #SQCR) AND "COG_FOLIE_L_is3800-Online" THEN #SQCR := #STEP_1010; END_IF;
END_REGION

REGION Network 11: INICIALIZACE 1015
   RUNG wire#powerrail
      { S7_Templates := "SrcType := Int" } EQ_Contact(in1 := #STEP_1010, in2 := #SQCR)
      Contact( "COG_FOLIE_P_is3800-Online" )
      Move(in := #STEP_1015, out1 => #SQCR)
   END_RUNG
   // the same network as SCL:
   IF (#STEP_1010 = #SQCR) AND "COG_FOLIE_P_is3800-Online" THEN #SQCR := #STEP_1015; END_IF;
END_REGION

REGION Network 12: INICIALIZACE 1020
   RUNG wire#powerrail
      { S7_Templates := "SrcType := Int" } EQ_Contact(in1 := #STEP_1015, in2 := #SQCR)
      Move(in := #STEP_5_HOME, out1 => #SQCR)
   END_RUNG
   // the same network as SCL:
   IF #STEP_1015 = #SQCR THEN #SQCR := #STEP_5_HOME; END_IF;
END_REGION

REGION Network 13: TRIGGER KAMER / automat control door
   RUNG wire#powerrail
      { S7_Templates := "SrcType := DInt" } LE_Contact(in1 := "DB_HMI_recype".VZDALENOST_KAMERA_ETIKETA_POZADOVANA, in2 := "DB_HMI_recype".aktualni_poloha)
      { S7_Templates := "SrcType := DInt" } NE_Contact(in1 := "DB_HMI_recype".aktualni_poloha, in2 := 0)
      { S7_Templates := "SrcType := DInt" } LT_Contact(in1 := "DB_HMI_recype".aktualni_poloha, in2 := 100)
      Coil( "COG_ETIKETA_COG_ETIKETA_is3800-Trigger" )
   END_RUNG
   RUNG wire#powerrail
      { S7_Templates := "SrcType := DInt" } LE_Contact(in1 := "DB_HMI_recype".VZDALENOST_KAMERY_FOLIE_POZADOVANA, in2 := "DB_HMI_recype".aktualni_poloha)
      { S7_Templates := "SrcType := DInt" } NE_Contact(in1 := "DB_HMI_recype".aktualni_poloha, in2 := 0)
      { S7_Templates := "SrcType := DInt" } LT_Contact(in1 := "DB_HMI_recype".aktualni_poloha, in2 := 180)
      wire#w1
      Coil( "COG_FOLIE_L_is3800-Trigger" )
   END_RUNG
   RUNG wire#w1
      Coil( "COG_FOLIE_P_is3800-Trigger" )
   END_RUNG
   // the same network as SCL:
   "COG_ETIKETA_COG_ETIKETA_is3800-Trigger" := ("DB_HMI_recype".VZDALENOST_KAMERA_ETIKETA_POZADOVANA <= "DB_HMI_recype".aktualni_poloha) AND ("DB_HMI_recype".aktualni_poloha <> 0) AND ("DB_HMI_recype".aktualni_poloha < 100);
   "COG_FOLIE_L_is3800-Trigger" := ("DB_HMI_recype".VZDALENOST_KAMERY_FOLIE_POZADOVANA <= "DB_HMI_recype".aktualni_poloha) AND ("DB_HMI_recype".aktualni_poloha <> 0) AND ("DB_HMI_recype".aktualni_poloha < 180);
   "COG_FOLIE_P_is3800-Trigger" := "COG_FOLIE_L_is3800-Trigger";
END_REGION

REGION Network 14: TRIGGER SVETEL
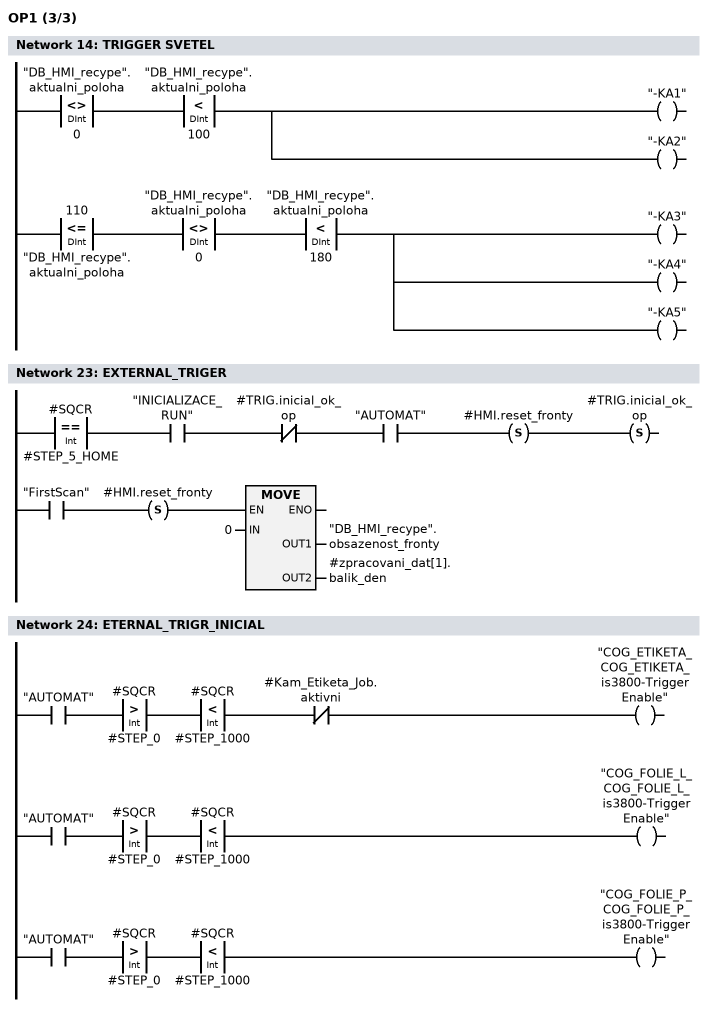
   RUNG wire#powerrail
      { S7_Templates := "SrcType := DInt" } NE_Contact(in1 := "DB_HMI_recype".aktualni_poloha, in2 := 0)
      { S7_Templates := "SrcType := DInt" } LT_Contact(in1 := "DB_HMI_recype".aktualni_poloha, in2 := 100)
      wire#w1
      Coil( "-KA1" )
   END_RUNG
   RUNG wire#w1
      Coil( "-KA2" )
   END_RUNG
   RUNG wire#powerrail
      { S7_Templates := "SrcType := DInt" } LE_Contact(in1 := 110, in2 := "DB_HMI_recype".aktualni_poloha)
      { S7_Templates := "SrcType := DInt" } NE_Contact(in1 := "DB_HMI_recype".aktualni_poloha, in2 := 0)
      { S7_Templates := "SrcType := DInt" } LT_Contact(in1 := "DB_HMI_recype".aktualni_poloha, in2 := 180)
      wire#w2
      Coil( "-KA3" )
   END_RUNG
   RUNG wire#w2
      Coil( "-KA4" )
   END_RUNG
   RUNG wire#w2
      Coil( "-KA5" )
   END_RUNG
   // the same network as SCL:
   "-KA1" := ("DB_HMI_recype".aktualni_poloha <> 0) AND ("DB_HMI_recype".aktualni_poloha < 100);
   "-KA2" := "-KA1";
   "-KA3" := (110 <= "DB_HMI_recype".aktualni_poloha) AND ("DB_HMI_recype".aktualni_poloha <> 0) AND ("DB_HMI_recype".aktualni_poloha < 180);
   "-KA4" := "-KA3";
   "-KA5" := "-KA3";
END_REGION

REGION Network 15 (SCL): TRIGGER MANUAL
   "iDB_CamManual"(xManEtiketa:="DB_Manual".xManEtiketa,
                   xManFolie:="DB_Manual".xManFolie);
END_REGION

REGION Network 16 (SCL): automat control data
   // Smyčka projde 104 bajtů (od 0 do 103)
   FOR #i := 0 TO 103 DO
       // PEEK čte přímo z paměti vstupů (16#81 = Periferní vstupy / Vstupy)
       // area 16#81 čte adresy %IB
       "DB_data_ctena".array_of_char[#i] := PEEK_BYTE(area := 16#81,
                                                       dbNumber := 0,
                                                       byteOffset := 76 + #i);
   END_FOR;

   // slozit text z prijatych znaku az po prvni $00
   "DB_data_ctena".upraveny := '';
   FOR #i := 0 TO 103 DO
       IF "DB_data_ctena".array_of_char[#i] = '$00' THEN
           EXIT;
       END_IF;
       "DB_data_ctena".upraveny := CONCAT(IN1 := "DB_data_ctena".upraveny,
                                          IN2 := CHAR_TO_STRING("DB_data_ctena".array_of_char[#i]));
   END_FOR;
END_REGION

REGION Network 17: automat control odfuk
END_REGION

REGION Network 18 (SCL): VYŘAZENÍ
   #Vyrazeni.s4_nabeh := #SENSORS.Pozice_vyrazovace AND NOT #Vyrazeni.s4_pamet;
   #Vyrazeni.s4_pamet := #SENSORS.Pozice_vyrazovace;

   IF "CONTROL_LINE_DB".trig.reset_error_all THEN
       #Vyrazeni.chyba_bez_dat := FALSE;
       #Vyrazeni.chyba_pist := FALSE;
       #Vyrazeni.alarm_nok_balik := FALSE;
   END_IF;

   IF NOT "AUTOMAT" THEN
       #Vyrazeni.aktivni := FALSE;
       #TIMER.TIMER_7.TON(IN := FALSE,
                          PT := #Vyrazeni.max_puls);
   ELSE
       REGION Plato prijelo k vyrazovaci - vzdy spotrebovat fronta[1]
           IF #Vyrazeni.s4_nabeh THEN
               IF "DB_HMI_recype".fronta[1].prenaseny_text = '' THEN
                   #Vyrazeni.chyba_bez_dat := TRUE;    // plato bez zaznamu ve fronte
                   #Vyrazeni.pocet_bez_dat := #Vyrazeni.pocet_bez_dat + 1;
                   #Vyrazeni.vyradit := TRUE;
               ELSE
                   #Vyrazeni.vyradit := "DB_HMI_recype".fronta[1].vyrazeni;
               END_IF;

               IF #Vyrazeni.vyradit THEN
                   #Vyrazeni.pocet_nok := #Vyrazeni.pocet_nok + 1;
                   IF "DB_HMI_recype".fronta[1].prenaseny_text = '' THEN
                       #Vyrazeni.posledni_nok_text := 'BEZ ZAZNAMU';
                       #Vyrazeni.posledni_nok_balik := 0;
                   ELSE
                       #Vyrazeni.posledni_nok_text := "DB_HMI_recype".fronta[1].prenaseny_text;
                       #Vyrazeni.posledni_nok_balik := "DB_HMI_recype".fronta[1].balik_den;
                   END_IF;
               END_IF;

               "DB_HMI_recype".fronta[1].prenaseny_text := '';
               "DB_HMI_recype".fronta[1].balik_den := 0;
               "DB_HMI_recype".fronta[1].vyrazeni := FALSE;

               IF #Vyrazeni.vyradit THEN
                   IF #Vyrazeni.vyrazovac_pripojen AND "DB_HMI_recype".recipe.vyrazovac_on_off THEN
                       #Vyrazeni.aktivni := TRUE;
                   ELSE
                       #Vyrazeni.alarm_nok_balik := TRUE;
                   END_IF;
               END_IF;
           END_IF;
       END_REGION

       REGION Pulz na vyrazovac - pevna delka Vyr.max_puls (200 ms)
           #TIMER.TIMER_7.TON(IN := #Vyrazeni.aktivni,
                              PT := #Vyrazeni.max_puls);
           IF #TIMER.TIMER_7.Q THEN
               #Vyrazeni.aktivni := FALSE;
           END_IF;
       END_REGION
   END_IF;

   // vystup na vyrazovac + rucni test (DB_Manual.test_vyr drzi vystup, dokud je TRUE)
   "RESERVE_DQ_2" := (#Vyrazeni.aktivni AND #Vyrazeni.vyrazovac_pripojen) OR "DB_Manual".test_vyr;

   // majak: po kazdem vyrazeni blika 5 s
   #Vyrazeni.majak_tp(IN := #Vyrazeni.aktivni AND #Vyrazeni.vyrazovac_pripojen,
                      PT := T#3S);
   #Vyrazeni.majak := #Vyrazeni.majak_tp.Q;
END_REGION

REGION Network 19 (SCL): CONTROL BLOCK presun_fronty
   IF "AUTOMAT" = true THEN


       REGION fronta 1 z 2
           IF "DB_HMI_recype".fronta[1].prenaseny_text = '' AND "DB_HMI_recype".fronta[2].prenaseny_text <> '' THEN
               "DB_HMI_recype".fronta[1]:= "DB_HMI_recype".fronta[2];
               "DB_HMI_recype".fronta[2].prenaseny_text := '';
               "DB_HMI_recype".fronta[2].balik_den := 0;
               "DB_HMI_recype".fronta[2].vyrazeni := false;
           END_IF;
       END_REGION

       REGION fronta 2 z 3
           IF "DB_HMI_recype".fronta[2].prenaseny_text = '' AND "DB_HMI_recype".fronta[3].prenaseny_text <> '' THEN
               "DB_HMI_recype".fronta[2] := "DB_HMI_recype".fronta[3];
               "DB_HMI_recype".fronta[3].prenaseny_text := '';
               "DB_HMI_recype".fronta[3].balik_den := 0;
               "DB_HMI_recype".fronta[3].vyrazeni := false;
           END_IF;
       END_REGION

       REGION fronta 3 z 4
           IF "DB_HMI_recype".fronta[3].prenaseny_text = '' AND "DB_HMI_recype".fronta[4].prenaseny_text <> '' THEN
               "DB_HMI_recype".fronta[3] := "DB_HMI_recype".fronta[4];
               "DB_HMI_recype".fronta[4].prenaseny_text := '';
               "DB_HMI_recype".fronta[4].balik_den := 0;
               "DB_HMI_recype".fronta[4].vyrazeni := false;
           END_IF;
       END_REGION

       REGION fronta 4 z 5
           IF "DB_HMI_recype".fronta[4].prenaseny_text = '' AND "DB_HMI_recype".fronta[5].prenaseny_text <> '' THEN
               "DB_HMI_recype".fronta[4] := "DB_HMI_recype".fronta[5];
               "DB_HMI_recype".fronta[5].prenaseny_text := '';
               "DB_HMI_recype".fronta[5].balik_den := 0;
               "DB_HMI_recype".fronta[5].vyrazeni := false;
           END_IF;
       END_REGION



   END_IF;


   REGION mazání fronty operátorem - bude pak možnost i automaticky ?
   IF #HMI.reset_fronty = true THEN

       "DB_HMI_recype".fronta[1].prenaseny_text := '';
       "DB_HMI_recype".fronta[1].balik_den := 0;
       "DB_HMI_recype".fronta[1].vyrazeni := false;

       "DB_HMI_recype".fronta[2].prenaseny_text := '';
       "DB_HMI_recype".fronta[2].balik_den := 0;
       "DB_HMI_recype".fronta[2].vyrazeni := false;

       "DB_HMI_recype".fronta[3].prenaseny_text := '';
       "DB_HMI_recype".fronta[3].balik_den := 0;
       "DB_HMI_recype".fronta[3].vyrazeni := false;

       "DB_HMI_recype".fronta[4].prenaseny_text := '';
       "DB_HMI_recype".fronta[4].balik_den := 0;
       "DB_HMI_recype".fronta[4].vyrazeni := false;

       "DB_HMI_recype".fronta[5].prenaseny_text := '';
       "DB_HMI_recype".fronta[5].balik_den := 0;
       "DB_HMI_recype".fronta[5].vyrazeni := false;

       "DB_HMI_recype".obsazenost_fronty := 0;
       #HMI.reset_fronty := false;

   END_IF;
   END_REGION;
END_REGION

REGION Network 20 (SCL)
   // ===== DENNI RESET POCITADLA PLAT (o pulnoci, lokalni cas) =====
   #ret := RD_LOC_T(#cas);
   IF #cas.HOUR = 0 AND #cas.MINUTE = 0 AND #cas.SECOND = 0 THEN
       #zpracovani_dat[1].balik_den := 0;
   END_IF;
   #aktual_kusy := #zpracovani_dat[1].balik_den;
END_REGION

REGION Network 21 (SCL): SBĚR VÝSLEDKŮ A ZÁPIS DO FRONTY
   #Kamera.s2_nabeh := #SENSORS.kontrola AND NOT #Kamera.s2_pamet;
   #Kamera.s2_pamet := #SENSORS.kontrola;

   IF NOT "AUTOMAT" THEN
       #Kamera.sber_aktivni := FALSE;
       #Kamera.last_id_etiketa := "COG_ETIKETA_is3800-InspectionID";
       #Kamera.last_id_folie_l := "COG_FOLIE_L_is3800-InspectionID";
       #Kamera.last_id_folie_p := "COG_FOLIE_P_is3800-InspectionID";
       #TIMER.TIMER_6.TON(IN := FALSE,
                          PT := #Kamera.timeout_sberu);
   ELSE
       REGION Prijem vysledku (zmena InspectionID = dokoncena inspekce)
           IF "COG_ETIKETA_is3800-InspectionID" <> #Kamera.last_id_etiketa THEN
               #Kamera.last_id_etiketa := "COG_ETIKETA_is3800-InspectionID";
               IF #Kamera.sber_aktivni THEN
                   #Kamera.prijato_etiketa := TRUE;
               END_IF;
           END_IF;
           // text prevzit, jakmile je k dispozici (i o par cyklu pozdeji nez ID);
           // prazdny vysledek dalsi inspekce dobry text neprepise
           IF #Kamera.sber_aktivni AND #Kamera.prijato_etiketa AND "DB_data_ctena".upraveny <> '' THEN
               #Kamera.text_etiketa := "DB_data_ctena".upraveny;
               #Kamera.ok_etiketa := TRUE;
           END_IF;
           IF "COG_FOLIE_L_is3800-InspectionID" <> #Kamera.last_id_folie_l THEN
               #Kamera.last_id_folie_l := "COG_FOLIE_L_is3800-InspectionID";
               IF #Kamera.sber_aktivni THEN
                   #Kamera.prijato_folie_l := TRUE;
                   #Kamera.ok_folie_l := ("COG_FOLIE_L_is3800-InspectionResults[0]" OR "COG_FOLIE_L_is3800-InspectionResults[1]") <> 16#00;
               END_IF;
           END_IF;
           IF "COG_FOLIE_P_is3800-InspectionID" <> #Kamera.last_id_folie_p THEN
               #Kamera.last_id_folie_p := "COG_FOLIE_P_is3800-InspectionID";
               IF #Kamera.sber_aktivni THEN
                   #Kamera.prijato_folie_p := TRUE;
                   #Kamera.ok_folie_p := ("COG_FOLIE_P_is3800-InspectionResults[0]" OR "COG_FOLIE_P_is3800-InspectionResults[1]") <> 16#00;
               END_IF;
           END_IF;
       END_REGION

       REGION Timeout - plato opustilo s2 a vysledky nedorazily
           #TIMER.TIMER_6.TON(IN := #Kamera.sber_aktivni AND NOT #SENSORS.kontrola,
                              PT := #Kamera.timeout_sberu);
       END_REGION

       REGION Vyhodnoceni a zapis do fronty
           IF #Kamera.sber_aktivni AND
               ((#Kamera.prijato_etiketa AND #Kamera.prijato_folie_l AND #Kamera.prijato_folie_p)
               OR #TIMER.TIMER_6.Q OR #Kamera.s2_nabeh) THEN

               #ocekavany_text := CONCAT(IN1 := "DB_HMI_recype".recipe.pole_string_2,
                                         IN2 := "DB_HMI_recype".recipe.pole_string_1);
               #format_etiketa_ok := #Kamera.bypass_ocr
               OR (FIND(IN1 := #Kamera.text_etiketa, IN2 := "DB_HMI_recype".recipe.pole_string_2) > 0
               AND NOT "OP2_DB".Tisk.datum_chyba);

               // kontrola kodu tridirny - nezavisla na bypass_ocr, vypinatelna z HMI
               #Kamera.tridirna_ok := NOT #Kamera.kontrola_tridirny
               OR FIND(IN1 := #Kamera.text_etiketa, IN2 := #KOD_TRIDIRNY) > 0;

               #Kamera.vyradit := NOT #Kamera.prijato_etiketa OR NOT #Kamera.prijato_folie_l
               OR NOT #Kamera.prijato_folie_p OR NOT #Kamera.ok_etiketa
               OR NOT #format_etiketa_ok OR NOT #Kamera.ok_folie_l
               OR NOT #Kamera.ok_folie_p
               OR NOT #Kamera.tridirna_ok;

